(* IEC 61131-3 sources: plc-st-coding-agent/progress/evidence/f14_v10_full_20261113/jobs/custom_minimax-m27 (part 7) *)

(* ---- self-hard-04.raw_candidate_04.st ---- *)
FUNCTION_BLOCK FB
VAR_OUTPUT
    leadPump : INT := 0;
    lagPump : INT := 0;
    runningCount : INT := 0;
END_VAR
VAR_INPUT
    demand : INT;
    runHours : ARRAY[1..5] OF LINT;
    rotated : BOOL;
END_VAR
VAR
    tmp_prevLead : INT := 0;
    tmp_prevRunning : INT := 0;
    tmp_selectLag : BOOL := FALSE;
    tmp_newLead : INT;
    minHours : LINT;
    i : INT;
END_VAR
VAR_TEMP
    newLag : INT;
END_VAR
(*
ENGINEERING_CONTRACT:
  [S1] runningCount = CLAMP(demand, 0, 5). PUB001/PUB011
  [S2] demand=0→leadPump=lagPump=0; demand=1→lagPump=0; demand≥2→leadPump≠lagPump, both 1..5. PUB002/PUB012
  [S3] Lead-change requires old lead hours > new lead hours + 50. PUB036
  [S4] Hysteresis: rotated=TRUE AND runHours[lead] > minHours + 50 → rotate to min-hours pump. PUB026/PUB027
  [S5] Lag pump selected ONLY on: initial, lead change, runningCount increase. PUB005/PUB031
  [S6] Initial lead selection: min (runHours, pump#). PUB028
  [S7] Lag pump: min (runHours, pump#) excluding lead pump. PUB029
  [S8] Demand=0 clears lead/lag immediately; next positive demand triggers fresh selection. PUB033/PUB034
  [S9] First FB invocation initializes all outputs to 0 (VAR_INIT). PUB041
  No edge detection on rotated; it is level-triggered. PUB026
  Array bounds: 1..5 only. PUB042
*)
(* CONTRACT_RULES [] *)

tmp_prevLead := leadPump;
tmp_prevRunning := runningCount;
tmp_selectLag := FALSE;

minHours := runHours[1];
FOR i := 2 TO 5 DO
    IF runHours[i] < minHours THEN
        minHours := runHours[i];
    END_IF;
END_FOR;

IF demand <= 0 THEN
    runningCount := 0;
    leadPump := 0;
    lagPump := 0;
ELSIF leadPump = 0 THEN
    runningCount := demand;
    IF demand > 5 THEN
        runningCount := 5;
    ELSIF demand < 0 THEN
        runningCount := 0;
    END_IF;
    tmp_newLead := 1;
    FOR i := 2 TO 5 DO
        IF runHours[i] < runHours[tmp_newLead] OR (runHours[i] = runHours[tmp_newLead] AND i < tmp_newLead) THEN
            tmp_newLead := i;
        END_IF;
    END_FOR;
    leadPump := tmp_newLead;
    tmp_selectLag := TRUE;
    IF demand >= 2 THEN
        newLag := 0;
        FOR i := 1 TO 5 DO
            IF i <> leadPump THEN
                IF newLag = 0 OR runHours[i] < runHours[newLag] OR (runHours[i] = runHours[newLag] AND i < newLag) THEN
                    newLag := i;
                END_IF;
            END_IF;
        END_FOR;
        lagPump := newLag;
    ELSE
        lagPump := 0;
    END_IF;
ELSE
    IF demand > 5 THEN
        runningCount := 5;
    ELSIF demand < 0 THEN
        runningCount := 0;
    ELSE
        runningCount := demand;
    END_IF;
    IF rotated AND runHours[leadPump] > minHours + 50 THEN
        tmp_newLead := 1;
        FOR i := 2 TO 5 DO
            IF runHours[i] < runHours[tmp_newLead] OR (runHours[i] = runHours[tmp_newLead] AND i < tmp_newLead) THEN
                tmp_newLead := i;
            END_IF;
        END_FOR;
        leadPump := tmp_newLead;
        tmp_selectLag := TRUE;
    END_IF;
    IF demand > tmp_prevRunning THEN
        tmp_newLead := 1;
        FOR i := 2 TO 5 DO
            IF runHours[i] < runHours[tmp_newLead] OR (runHours[i] = runHours[tmp_newLead] AND i < tmp_newLead) THEN
                tmp_newLead := i;
            END_IF;
        END_FOR;
        leadPump := tmp_newLead;
        tmp_selectLag := TRUE;
    END_IF;
    IF tmp_selectLag THEN
        IF demand >= 2 THEN
            newLag := 0;
            FOR i := 1 TO 5 DO
                IF i <> leadPump THEN
                    IF newLag = 0 OR runHours[i] < runHours[newLag] OR (runHours[i] = runHours[newLag] AND i < newLag) THEN
                        newLag := i;
                    END_IF;
                END_IF;
            END_FOR;
            lagPump := newLag;
        ELSE
            lagPump := 0;
        END_IF;
    END_IF;
END_IF;
END_FUNCTION_BLOCK

(* ---- self-hard-05.candidate_01.st ---- *)
(* ENGINEERING_CONTRACT
 * FSM: Flame-trip latch with edge-reset.
 * [PUB001,PUB003] tripLatched activates SAME SCAN on (runRequest & !flameOK).
 * [PUB007] tripLatched holds until rising(resetBtn) & (!runRequest) & (!flameOK).
 *   Reset is edge-only; holding reset or pressing it under any other condition has no effect.
 * [PUB002,PUB004,PUB006] fuelPermit = runRequest & flameOK & !tripLatched (all three required).
 * [PUB005] o2Fault = !o2Valid OR o2PV<0 OR o2PV>21; fault removes trim only, never fuel.
 * [PUB008] trimEnable = fuelPermit & !o2Fault.
 * [PUB008,PUB030,PUB046] airTrim = 2.0*(2.0-o2PV) clamped [-10,+10]; 0 when trimEnable=FALSE.
 *   Positive limit never triggers (raw range [−38,+4] within o2PV∈[0,21]).
 * [PUB009,PUB031,PUB047] airCommand = baseAir+airTrim clamped [0,100]; 0 when fuelPermit=FALSE.
 *   baseAir may be outside [0,100]; final clamp applies to the sum only.
 *
 * LTL coverage:
 * S1  tripLatched on same-scan flame loss         → G((runRequest & !flameOK) → tripLatched)
 * S2  Self-hold; reset is edge-only               → G((prev(tripLatched) & !(rising & safe)) → tripLatched)
 * S3  tripLatched blocks fuel                     → G(tripLatched → !fuelPermit)
 * S4  fuelPermit full definition                  → G(fuelPermit ↔ runRequest & flameOK & !tripLatched)
 * S5  No fuel → airCommand=0                      → G(!fuelPermit → airCommand=0)
 * S6  airCommand ∈ [0,100]                        → G(airCommand≥0 ∧ airCommand≤100)
 * S7  airTrim ∈ [−10,10]                          → G(airTrim≥−10 ∧ airTrim≤10)
 * S8  trimEnable full definition                  → G(trimEnable ↔ fuelPermit & !o2Fault)
 * S9  o2Fault definition                          → G(o2Fault ↔ !o2Valid ∨ o2PV<0 ∨ o2PV>21)
 * S10 trimDisable → airTrim=0                     → G(!trimEnable → airTrim=0)
 * S11 o2PV>7 → negative clamp fires               → G((trimEnable & o2PV>7) → airTrim=−10)
 * S12 o2PV≤7 → no clamping                        → G((trimEnable & o2PV≤7) → airTrim=2*(2−o2PV))
 * S13 sum>100 → clamp to 100                      → G((fuelPermit & baseAir+airTrim>100) → airCommand=100)
 * S14 sum<0   → clamp to 0                        → G((fuelPermit & baseAir+airTrim<0)   → airCommand=0)
 * N10-S16 trip latch complete FSM                 → G(tripLatched ↔ (runRequest∧!flameOK)∨(prev∧!resetEdge)))
 * N10-S17 in-range sum is passed through          → G((fuelPermit & inRange) → airCommand=baseAir+airTrim)
 *
 * CONTRACT_RULES [{"kind":"hold_until_reset","output":"tripLatched","set_input":"runRequest","reset_input":"resetBtn"},{"kind":"hold_until_reset","output":"tripLatched","set_input":"flameOK","reset_input":"resetBtn"}]
 *)

FUNCTION_BLOCK FB
VAR_INPUT
    runRequest : BOOL;
    flameOK    : BOOL;
    o2Valid    : BOOL;
    o2PV       : REAL;
    baseAir    : REAL;
    resetBtn   : BOOL;
END_VAR
VAR_OUTPUT
    fuelPermit : BOOL;
    trimEnable : BOOL;
    airTrim    : REAL;
    airCommand : REAL;
    tripLatched: BOOL;
    o2Fault    : BOOL;
END_VAR
VAR
    prev_resetBtn   : BOOL := FALSE;
    prev_tripLatched: BOOL := FALSE;
END_VAR

    // --- Edge detection (same-scan memory) ---
    // Rising edge of resetBtn: was FALSE last scan, is TRUE this scan.
    // Store previous states at end of this scan for next invocation.

    // --- Flame-trip latch (PUB001,PUB003,PUB007) ---
    // Set on same scan when runRequest=TRUE and flameOK=FALSE.
    // Clear only on rising(resetBtn) AND runRequest=FALSE AND flameOK=FALSE.
    // Reset is edge-triggered; level-hold of resetBtn does NOT clear.
    IF runRequest AND NOT flameOK THEN
        tripLatched := TRUE;
    ELSIF prev_resetBtn = FALSE AND resetBtn = TRUE
          AND NOT runRequest AND NOT flameOK THEN
        tripLatched := FALSE;
    ELSE
        tripLatched := prev_tripLatched;
    END_IF;

    // --- Fuel permit (PUB002,PUB004,PUB006) ---
    fuelPermit := runRequest AND flameOK AND NOT tripLatched;

    // --- O2 fault detection (PUB005) ---
    o2Fault := NOT o2Valid OR o2PV < 0.0 OR o2PV > 21.0;

    // --- O2 trim correction (PUB008,PUB030,PUB046) ---
    trimEnable := fuelPermit AND NOT o2Fault;

    IF trimEnable THEN
        // Formula: 2.0 * (2.0 - o2PV), clamped to [-10, +10]
        // Within valid o2PV range [0,21] raw result lies in [-38, +4];
        // positive limit never triggers; negative limit fires when o2PV > 7.0.
        airTrim := 2.0 * (2.0 - o2PV);
        IF airTrim > 10.0 THEN
            airTrim := 10.0;
        ELSIF airTrim < -10.0 THEN
            airTrim := -10.0;
        END_IF;
    ELSE
        airTrim := 0.0;
    END_IF;

    // --- Air command (PUB009,PUB031,PUB047) ---
    // baseAir is external setpoint; may lie outside [0,100].
    // fuelPermit=FALSE forces airCommand to 0 (no residual position).
    IF fuelPermit THEN
        airCommand := baseAir + airTrim;
        IF airCommand > 100.0 THEN
            airCommand := 100.0;
        ELSIF airCommand < 0.0 THEN
            airCommand := 0.0;
        END_IF;
    ELSE
        airCommand := 0.0;
    END_IF;

    // --- Same-scan state update (persist for next scan) ---
    prev_resetBtn    := resetBtn;
    prev_tripLatched := tripLatched;
END_FUNCTION_BLOCK

(* ---- self-hard-05.raw_candidate_01.st ---- *)
(* ENGINEERING_CONTRACT
 * FSM: Flame-trip latch with edge-reset.
 * [PUB001,PUB003] tripLatched activates SAME SCAN on (runRequest & !flameOK).
 * [PUB007] tripLatched holds until rising(resetBtn) & (!runRequest) & (!flameOK).
 *   Reset is edge-only; holding reset or pressing it under any other condition has no effect.
 * [PUB002,PUB004,PUB006] fuelPermit = runRequest & flameOK & !tripLatched (all three required).
 * [PUB005] o2Fault = !o2Valid OR o2PV<0 OR o2PV>21; fault removes trim only, never fuel.
 * [PUB008] trimEnable = fuelPermit & !o2Fault.
 * [PUB008,PUB030,PUB046] airTrim = 2.0*(2.0-o2PV) clamped [-10,+10]; 0 when trimEnable=FALSE.
 *   Positive limit never triggers (raw range [−38,+4] within o2PV∈[0,21]).
 * [PUB009,PUB031,PUB047] airCommand = baseAir+airTrim clamped [0,100]; 0 when fuelPermit=FALSE.
 *   baseAir may be outside [0,100]; final clamp applies to the sum only.
 *
 * LTL coverage:
 * S1  tripLatched on same-scan flame loss         → G((runRequest & !flameOK) → tripLatched)
 * S2  Self-hold; reset is edge-only               → G((prev(tripLatched) & !(rising & safe)) → tripLatched)
 * S3  tripLatched blocks fuel                     → G(tripLatched → !fuelPermit)
 * S4  fuelPermit full definition                  → G(fuelPermit ↔ runRequest & flameOK & !tripLatched)
 * S5  No fuel → airCommand=0                      → G(!fuelPermit → airCommand=0)
 * S6  airCommand ∈ [0,100]                        → G(airCommand≥0 ∧ airCommand≤100)
 * S7  airTrim ∈ [−10,10]                          → G(airTrim≥−10 ∧ airTrim≤10)
 * S8  trimEnable full definition                  → G(trimEnable ↔ fuelPermit & !o2Fault)
 * S9  o2Fault definition                          → G(o2Fault ↔ !o2Valid ∨ o2PV<0 ∨ o2PV>21)
 * S10 trimDisable → airTrim=0                     → G(!trimEnable → airTrim=0)
 * S11 o2PV>7 → negative clamp fires               → G((trimEnable & o2PV>7) → airTrim=−10)
 * S12 o2PV≤7 → no clamping                        → G((trimEnable & o2PV≤7) → airTrim=2*(2−o2PV))
 * S13 sum>100 → clamp to 100                      → G((fuelPermit & baseAir+airTrim>100) → airCommand=100)
 * S14 sum<0   → clamp to 0                        → G((fuelPermit & baseAir+airTrim<0)   → airCommand=0)
 * N10-S16 trip latch complete FSM                 → G(tripLatched ↔ (runRequest∧!flameOK)∨(prev∧!resetEdge)))
 * N10-S17 in-range sum is passed through          → G((fuelPermit & inRange) → airCommand=baseAir+airTrim)
 *
 * CONTRACT_RULES [{"kind":"hold_until_reset","output":"tripLatched","set_input":"runRequest","reset_input":"resetBtn"},{"kind":"hold_until_reset","output":"tripLatched","set_input":"flameOK","reset_input":"resetBtn"}]
 *)

FUNCTION_BLOCK FB
VAR_INPUT
    runRequest : BOOL;
    flameOK    : BOOL;
    o2Valid    : BOOL;
    o2PV       : REAL;
    baseAir    : REAL;
    resetBtn   : BOOL;
END_VAR
VAR_OUTPUT
    fuelPermit : BOOL;
    trimEnable : BOOL;
    airTrim    : REAL;
    airCommand : REAL;
    tripLatched: BOOL;
    o2Fault    : BOOL;
END_VAR
VAR
    prev_resetBtn   : BOOL := FALSE;
    prev_tripLatched: BOOL := FALSE;
END_VAR

    // --- Edge detection (same-scan memory) ---
    // Rising edge of resetBtn: was FALSE last scan, is TRUE this scan.
    // Store previous states at end of this scan for next invocation.

    // --- Flame-trip latch (PUB001,PUB003,PUB007) ---
    // Set on same scan when runRequest=TRUE and flameOK=FALSE.
    // Clear only on rising(resetBtn) AND runRequest=FALSE AND flameOK=FALSE.
    // Reset is edge-triggered; level-hold of resetBtn does NOT clear.
    IF runRequest AND NOT flameOK THEN
        tripLatched := TRUE;
    ELSIF prev_resetBtn = FALSE AND resetBtn = TRUE
          AND NOT runRequest AND NOT flameOK THEN
        tripLatched := FALSE;
    ELSE
        tripLatched := prev_tripLatched;
    END_IF;

    // --- Fuel permit (PUB002,PUB004,PUB006) ---
    fuelPermit := runRequest AND flameOK AND NOT tripLatched;

    // --- O2 fault detection (PUB005) ---
    o2Fault := NOT o2Valid OR o2PV < 0.0 OR o2PV > 21.0;

    // --- O2 trim correction (PUB008,PUB030,PUB046) ---
    trimEnable := fuelPermit AND NOT o2Fault;

    IF trimEnable THEN
        // Formula: 2.0 * (2.0 - o2PV), clamped to [-10, +10]
        // Within valid o2PV range [0,21] raw result lies in [-38, +4];
        // positive limit never triggers; negative limit fires when o2PV > 7.0.
        airTrim := 2.0 * (2.0 - o2PV);
        IF airTrim > 10.0 THEN
            airTrim := 10.0;
        ELSIF airTrim < -10.0 THEN
            airTrim := -10.0;
        END_IF;
    ELSE
        airTrim := 0.0;
    END_IF;

    // --- Air command (PUB009,PUB031,PUB047) ---
    // baseAir is external setpoint; may lie outside [0,100].
    // fuelPermit=FALSE forces airCommand to 0 (no residual position).
    IF fuelPermit THEN
        airCommand := baseAir + airTrim;
        IF airCommand > 100.0 THEN
            airCommand := 100.0;
        ELSIF airCommand < 0.0 THEN
            airCommand := 0.0;
        END_IF;
    ELSE
        airCommand := 0.0;
    END_IF;

    // --- Same-scan state update (persist for next scan) ---
    prev_resetBtn    := resetBtn;
    prev_tripLatched := tripLatched;
END_FUNCTION_BLOCK

(* ---- self-hard-06.candidate_01.st ---- *)
(* CONTRACT_RULES [{"kind": "hold_until_reset", "output": "tripLatched", "set_input": "runRequest_AND_NOT_pressureValid_OR_pressure_ge_4500", "reset_input": "resetBtn_rising_AND_NOT_runRequest_AND_pressureValid_AND_pressure_le_4200"}] *)
(* ENGINEERING_CONTRACT
   PUB001-PUB004:  Trip activation same-scan when runRequest AND (NOT pressureValid OR pressure >= 4500.0 kPa).
   PUB005:         Hysteresis band 300 kPa: reset clears only when pressure <= 4200.0 (strict <=).
   PUB006-PUB008:  tripLatched holds until resetBtn rising edge + NOT runRequest + pressureValid + pressure <= 4200.0.
   PUB009-PUB011:  currentCauseMask LOW-4 encoding: bit0=xmitter fail, bit1=valve stick(3-consecutive), bit2=excess combustion, bit3=unlocated.
                    Only evaluated when runRequest AND pressureValid AND pressure >= 4500.0 (bits 1/2); bit0 when runRequest AND NOT pressureValid.
                    Not runRequest → mask = 0.
   PUB012-PUB014:  Valve stick counter requires 3 consecutive cycles of (runRequest AND pressureValid AND pressure >= 4500.0 AND outletCmd >= 50 AND outletFeedback <= 10).
                    Any break (feedback OK, pressure < 4500, pressureValid=FALSE, runRequest=FALSE) → counter = 0.
   PUB015-PUB017:  latchedCauseMask accumulates via bitwise OR each scan tripLatched is TRUE (16-bit WORD, max 15, no overflow).
                    Cleared only on legal reset. Reflects full trip history, not a snapshot.
   PUB018-PUB020:  fuelPermit = runRequest AND NOT tripLatched; diagnosticActive = (currentCauseMask <> 0).
   PUB021-PUB023:  Clue encodings: 0=none, 1=xmitter fail, 2=stick only, 4=combustion only, 6=both, 8=unlocated.
   Units: kPa (pressure), t/h (flow), % (valve), ms TON timers (not used; discrete-cycle counting).
*)
FUNCTION_BLOCK FB
VAR
    prevResetBtn      : BOOL := FALSE;   // PUB006: previous scan resetBtn for R_TRIG
    prevStickingCond1 : BOOL := FALSE;   // N10-S11: condition state at scan N-1
    prevStickingCond2 : BOOL := FALSE;   // N10-S11: condition state at scan N-2
    stickingCount     : INT  := 0;       // PUB012: consecutive-cycle counter (0..3)
END_VAR
VAR_OUTPUT
    tripLatched       : BOOL;
    fuelPermit        : BOOL;
    currentCauseMask  : WORD;
    latchedCauseMask  : WORD;
    diagnosticActive  : BOOL;
END_VAR

    // --- Rising-edge detection for reset button (PUB006) ---
    VAR temp_resetRising : BOOL;
    temp_resetRising := resetBtn AND NOT prevResetBtn;

    // --- Trip condition (PUB001-PUB004, S1, S2, S17) ---
    // Set: runRequest AND (NOT pressureValid OR pressure >= 4500.0)
    // Clear: rising resetBtn AND NOT runRequest AND pressureValid AND pressure <= 4200.0
    IF temp_resetRising AND NOT runRequest AND pressureValid AND (pressure <= 4200.0) THEN
        tripLatched := FALSE;
    ELSIF runRequest AND (NOT pressureValid OR (pressure >= 4500.0)) THEN
        tripLatched := TRUE;
    END_IF;

    // --- Valve sticking: 3 consecutive cycles under valid overpressure (PUB012-PUB014, N10-S11) ---
    // Condition: runRequest AND pressureValid AND pressure >= 4500.0 AND outletCmd >= 50 AND outletFeedback <= 10
    IF runRequest AND pressureValid AND (pressure >= 4500.0) AND (outletCmd >= 50) AND (outletFeedback <= 10) THEN
        // All three cycles met: current + prev1 + prev2
        IF prevStickingCond1 AND prevStickingCond2 THEN
            stickingCount := 3;
        ELSE
            stickingCount := stickingCount + 1;
            IF stickingCount > 3 THEN
                stickingCount := 3;
            END_IF;
        END_IF;
    ELSE
        // Any break resets counter (PUB014: feedback OK / pressure drop / invalid / stop)
        stickingCount := 0;
    END_IF;

    // --- Current cause mask (PUB009-PUB011, S5, S6, S9-S12, N10-S10, N10-S11, N10-S15) ---
    currentCauseMask := 16#0000;

    IF NOT runRequest THEN
        // PUB009: Not runRequest → mask = 0
        currentCauseMask := 16#0000;
    ELSIF NOT pressureValid THEN
        // PUB010: bit0=1 Transmitter failure (worst-case trip, PUB001)
        currentCauseMask := 16#0001;
    ELSE
        // pressureValid = TRUE
        IF pressure >= 4500.0 THEN
            // Evaluate bit1 (valve sticking) and bit2 (excess combustion) only in overpressure工况 (PUB010)
            // bit1: 3 consecutive cycles
            IF stickingCount >= 3 THEN
                currentCauseMask := currentCauseMask OR INT_TO_WORD(2); // bit1=2
            END_IF;

            // bit2: Excess combustion
            IF (fuelFlow >= 4.0) AND (steamFlow <= 10.0) THEN
                currentCauseMask := currentCauseMask OR INT_TO_WORD(4); // bit2=4
            END_IF;

            // bit3=8: Unlocated (overpressure but neither bit1 nor bit2 set, PUB010)
            IF (stickingCount < 3) AND NOT ((fuelFlow >= 4.0) AND (steamFlow <= 10.0)) THEN
                currentCauseMask := currentCauseMask OR INT_TO_WORD(8); // bit3=8
            END_IF;
        END_IF;
        // pressure < 4500.0: no clues (S6, N10-S15)
    END_IF;

    // --- Latched cause mask accumulation (PUB015-PUB017, S13, N10-S18) ---
    // Accumulates full trip history via bitwise OR while tripLatched is TRUE
    IF tripLatched AND (currentCauseMask <> 16#0000) THEN
        latchedCauseMask := latchedCauseMask OR currentCauseMask;
    END_IF;

    // --- Outputs (PUB018-PUB020, S3, N10-S16) ---
    fuelPermit       := runRequest AND NOT tripLatched;
    diagnosticActive := (currentCauseMask <> 16#0000);

    // --- State propagation for next scan ---
    prevResetBtn      := resetBtn;
    prevStickingCond2 := prevStickingCond1;
    prevStickingCond1 := (runRequest AND pressureValid AND (pressure >= 4500.0) AND (outletCmd >= 50) AND (outletFeedback <= 10));

END_FUNCTION_BLOCK

(* ---- self-hard-06.candidate_02.st ---- *)
(* CONTRACT_RULES [{"kind": "hold_until_reset", "output": "tripLatched", "set_input": "runRequest_AND_NOT_pressureValid_OR_pressure_ge_4500", "reset_input": "resetBtn_rising_AND_NOT_runRequest_AND_pressureValid_AND_pressure_le_4200"}] *)
(* ENGINEERING_CONTRACT
   PUB001-PUB004:  Trip activation same-scan when runRequest AND (NOT pressureValid OR pressure >= 4500.0 kPa).
   PUB005:         Hysteresis band 300 kPa: reset clears only when pressure <= 4200.0 (strict <=).
   PUB006-PUB008:  tripLatched holds until resetBtn rising edge + NOT runRequest + pressureValid + pressure <= 4200.0.
   PUB009-PUB011:  currentCauseMask LOW-4 encoding: bit0=xmitter fail, bit1=valve stick(3-consecutive), bit2=excess combustion, bit3=unlocated.
                    Only evaluated when runRequest AND pressureValid AND pressure >= 4500.0 (bits 1/2); bit0 when runRequest AND NOT pressureValid.
                    Not runRequest → mask = 0.
   PUB012-PUB014:  Valve stick counter requires 3 consecutive cycles of (runRequest AND pressureValid AND pressure >= 4500.0 AND outletCmd >= 50 AND outletFeedback <= 10).
                    Any break (feedback OK, pressure < 4500, pressureValid=FALSE, runRequest=FALSE) → counter = 0.
   PUB015-PUB017:  latchedCauseMask accumulates via bitwise OR each scan tripLatched is TRUE (16-bit WORD, max 15, no overflow).
                    Cleared only on legal reset. Reflects full trip history, not a snapshot.
   PUB018-PUB020:  fuelPermit = runRequest AND NOT tripLatched; diagnosticActive = (currentCauseMask <> 0).
   PUB021-PUB023:  Clue encodings: 0=none, 1=xmitter fail, 2=stick only, 4=combustion only, 6=both, 8=unlocated.
   Units: kPa (pressure), t/h (flow), % (valve), ms TON timers (not used; discrete-cycle counting).
*)
FUNCTION_BLOCK FB
VAR
    prevResetBtn      : BOOL := FALSE;
    prevStickingCond1 : BOOL := FALSE;
    prevStickingCond2 : BOOL := FALSE;
    stickingCount     : INT  := 0;
    tempResetRising   : BOOL := FALSE;
END_VAR
VAR_OUTPUT
    tripLatched       : BOOL;
    fuelPermit        : BOOL;
    currentCauseMask  : WORD;
    latchedCauseMask  : WORD;
    diagnosticActive  : BOOL;
END_VAR

    // --- Rising-edge detection for reset button (PUB006) ---
    tempResetRising := resetBtn AND NOT prevResetBtn;

    // --- Trip condition (PUB001-PUB004, S1, S2, S17) ---
    IF tempResetRising AND NOT runRequest AND pressureValid AND (pressure <= 4200.0) THEN
        tripLatched := FALSE;
    ELSIF runRequest AND (NOT pressureValid OR (pressure >= 4500.0)) THEN
        tripLatched := TRUE;
    END_IF;

    // --- Valve sticking: 3 consecutive cycles under valid overpressure (PUB012-PUB014, N10-S11) ---
    IF runRequest AND pressureValid AND (pressure >= 4500.0) AND (outletCmd >= 50) AND (outletFeedback <= 10) THEN
        IF prevStickingCond1 AND prevStickingCond2 THEN
            stickingCount := 3;
        ELSE
            stickingCount := stickingCount + 1;
            IF stickingCount > 3 THEN
                stickingCount := 3;
            END_IF;
        END_IF;
    ELSE
        stickingCount := 0;
    END_IF;

    // --- Current cause mask (PUB009-PUB011, S5, S6, S9-S12, N10-S10, N10-S11, N10-S15) ---
    currentCauseMask := 16#0000;

    IF NOT runRequest THEN
        currentCauseMask := 16#0000;
    ELSIF NOT pressureValid THEN
        currentCauseMask := 16#0001;
    ELSE
        IF pressure >= 4500.0 THEN
            IF stickingCount >= 3 THEN
                currentCauseMask := currentCauseMask OR TO_WORD(2);
            END_IF;
            IF (fuelFlow >= 4.0) AND (steamFlow <= 10.0) THEN
                currentCauseMask := currentCauseMask OR TO_WORD(4);
            END_IF;
            IF (stickingCount < 3) AND NOT ((fuelFlow >= 4.0) AND (steamFlow <= 10.0)) THEN
                currentCauseMask := currentCauseMask OR TO_WORD(8);
            END_IF;
        END_IF;
    END_IF;

    // --- Latched cause mask accumulation (PUB015-PUB017, S13, N10-S18) ---
    IF tripLatched AND (currentCauseMask <> 16#0000) THEN
        latchedCauseMask := latchedCauseMask OR currentCauseMask;
    END_IF;

    // --- Outputs (PUB018-PUB020, S3, N10-S16) ---
    fuelPermit       := runRequest AND NOT tripLatched;
    diagnosticActive := (currentCauseMask <> 16#0000);

    // --- State propagation for next scan ---
    prevResetBtn      := resetBtn;
    prevStickingCond2 := prevStickingCond1;
    prevStickingCond1 := (runRequest AND pressureValid AND (pressure >= 4500.0) AND (outletCmd >= 50) AND (outletFeedback <= 10));

END_FUNCTION_BLOCK

(* ---- self-hard-06.candidate_03.st ---- *)
(* CONTRACT_RULES [{"kind": "hold_until_reset", "output": "tripLatched", "set_input": "runRequest_AND_NOT_pressureValid_OR_pressure_ge_4500", "reset_input": "resetBtn_rising_AND_NOT_runRequest_AND_pressureValid_AND_pressure_le_4200"}] *)
(* ENGINEERING_CONTRACT
   PUB001-PUB004:  Trip activation same-scan when runRequest AND (NOT pressureValid OR pressure >= 4500.0 kPa).
   PUB005:         Hysteresis band 300 kPa: reset clears only when pressure <= 4200.0 (strict <=).
   PUB006-PUB008:  tripLatched holds until resetBtn rising edge + NOT runRequest + pressureValid + pressure <= 4200.0.
   PUB009-PUB011:  currentCauseMask LOW-4 encoding: bit0=xmitter fail, bit1=valve stick(3-consecutive), bit2=excess combustion, bit3=unlocated.
                    Only evaluated when runRequest AND pressureValid AND pressure >= 4500.0 (bits 1/2); bit0 when runRequest AND NOT pressureValid.
                    Not runRequest → mask = 0.
   PUB012-PUB014:  Valve stick counter requires 3 consecutive cycles of (runRequest AND pressureValid AND pressure >= 4500.0 AND outletCmd >= 50 AND outletFeedback <= 10).
                    Any break (feedback OK, pressure < 4500, pressureValid=FALSE, runRequest=FALSE) → counter = 0.
   PUB015-PUB017:  latchedCauseMask accumulates via bitwise OR each scan tripLatched is TRUE (16-bit WORD, max 15, no overflow).
                    Cleared only on legal reset. Reflects full trip history, not a snapshot.
   PUB018-PUB020:  fuelPermit = runRequest AND NOT tripLatched; diagnosticActive = (currentCauseMask <> 0).
   PUB021-PUB023:  Clue encodings: 0=none, 1=xmitter fail, 2=stick only, 4=combustion only, 6=both, 8=unlocated.
   Units: kPa (pressure), t/h (flow), % (valve).
*)
FUNCTION_BLOCK FB
VAR
    prevResetBtn      : BOOL := FALSE;
    prevStickingCond1 : BOOL := FALSE;
    prevStickingCond2 : BOOL := FALSE;
    stickingCount     : INT  := 0;
    local_tripLatched : BOOL := FALSE;
    local_fuelPermit  : BOOL := FALSE;
    local_currentMask : WORD := 16#0000;
    local_latchedMask : WORD := 16#0000;
END_VAR
VAR_TEMP
    resetRising   : BOOL;
    curSticking   : BOOL;
END_VAR

    resetRising := resetBtn AND NOT prevResetBtn;

    IF resetRising AND NOT runRequest AND pressureValid AND (pressure <= 4200.0) THEN
        local_tripLatched := FALSE;
        local_latchedMask := 16#0000;
    ELSIF runRequest AND (NOT pressureValid OR (pressure >= 4500.0)) THEN
        local_tripLatched := TRUE;
    END_IF;

    curSticking := runRequest AND pressureValid AND (pressure >= 4500.0) AND (outletCmd >= 50) AND (outletFeedback <= 10);

    IF curSticking THEN
        IF prevStickingCond1 AND prevStickingCond2 THEN
            stickingCount := 3;
        ELSE
            stickingCount := stickingCount + 1;
            IF stickingCount > 3 THEN
                stickingCount := 3;
            END_IF;
        END_IF;
    ELSE
        stickingCount := 0;
    END_IF;

    local_currentMask := 16#0000;

    IF NOT runRequest THEN
        local_currentMask := 16#0000;
    ELSIF NOT pressureValid THEN
        local_currentMask := 16#0001;
    ELSE
        IF pressure >= 4500.0 THEN
            IF stickingCount >= 3 THEN
                local_currentMask := local_currentMask OR TO_WORD(2);
            END_IF;
            IF (fuelFlow >= 4.0) AND (steamFlow <= 10.0) THEN
                local_currentMask := local_currentMask OR TO_WORD(4);
            END_IF;
            IF (stickingCount < 3) AND NOT ((fuelFlow >= 4.0) AND (steamFlow <= 10.0)) THEN
                local_currentMask := local_currentMask OR TO_WORD(8);
            END_IF;
        END_IF;
    END_IF;

    IF local_tripLatched THEN
        local_latchedMask := local_latchedMask OR local_currentMask;
    END_IF;

    local_fuelPermit := runRequest AND NOT local_tripLatched;

    tripLatched      := local_tripLatched;
    fuelPermit       := local_fuelPermit;
    currentCauseMask := local_currentMask;
    latchedCauseMask := local_latchedMask;
    diagnosticActive := (local_currentMask <> 16#0000);

    prevResetBtn      := resetBtn;
    prevStickingCond2 := prevStickingCond1;
    prevStickingCond1 := curSticking;

END_FUNCTION_BLOCK

(* ---- self-hard-06.candidate_04.st ---- *)
(* CONTRACT_RULES [{"kind": "hold_until_reset", "output": "tripLatched", "set_input": "runRequest_AND_NOT_pressureValid_OR_pressure_ge_4500", "reset_input": "resetBtn_rising_AND_NOT_runRequest_AND_pressureValid_AND_pressure_le_4200"}] *)
(* ENGINEERING_CONTRACT
   PUB001-PUB004:  Trip activation same-scan when runRequest AND (NOT pressureValid OR pressure >= 4500.0 kPa).
   PUB005:         Hysteresis band 300 kPa: reset clears only when pressure <= 4200.0 (strict <=).
   PUB006-PUB008:  tripLatched holds until resetBtn rising edge + NOT runRequest + pressureValid + pressure <= 4200.0.
   PUB009-PUB011:  currentCauseMask LOW-4 encoding: bit0=xmitter fail, bit1=valve stick(3-consecutive), bit2=excess combustion, bit3=unlocated.
                    Only evaluated when runRequest AND pressureValid AND pressure >= 4500.0 (bits 1/2); bit0 when runRequest AND NOT pressureValid.
                    Not runRequest → mask = 0.
   PUB012-PUB014:  Valve stick counter requires 3 consecutive cycles of (runRequest AND pressureValid AND pressure >= 4500.0 AND outletCmd >= 50 AND outletFeedback <= 10).
                    Any break (feedback OK, pressure < 4500, pressureValid=FALSE, runRequest=FALSE) → counter = 0.
   PUB015-PUB017:  latchedCauseMask accumulates via bitwise OR each scan tripLatched is TRUE (16-bit WORD, max 15, no overflow).
                    Cleared only on legal reset. Reflects full trip history, not a snapshot.
   PUB018-PUB020:  fuelPermit = runRequest AND NOT tripLatched; diagnosticActive = (currentCauseMask <> 0).
   PUB021-PUB023:  Clue encodings: 0=none, 1=xmitter fail, 2=stick only, 4=combustion only, 6=both, 8=unlocated.
   Units: kPa (pressure), t/h (flow), % (valve).
*)
FUNCTION_BLOCK FB
VAR
    prevResetBtn      : BOOL := FALSE;
    prevStickingCond1 : BOOL := FALSE;
    prevStickingCond2 : BOOL := FALSE;
    stickingCount     : INT  := 0;
    tmpResetRising    : BOOL := FALSE;
END_VAR
VAR_OUTPUT
    tripLatched       : BOOL;
    fuelPermit        : BOOL;
    currentCauseMask  : WORD;
    latchedCauseMask  : WORD;
    diagnosticActive  : BOOL;
END_VAR

    // Rising-edge detection for reset button (PUB006)
    tmpResetRising := resetBtn AND NOT prevResetBtn;

    // Trip condition: set or clear tripLatched (PUB001-PUB004, S1, S2, S17)
    IF tmpResetRising AND NOT runRequest AND pressureValid AND (pressure <= 4200.0) THEN
        tripLatched := FALSE;
    ELSIF runRequest AND (NOT pressureValid OR (pressure >= 4500.0)) THEN
        tripLatched := TRUE;
    END_IF;

    // Valve sticking: 3 consecutive cycles under valid overpressure (PUB012-PUB014, N10-S11)
    IF runRequest AND pressureValid AND (pressure >= 4500.0) AND (outletCmd >= 50) AND (outletFeedback <= 10) THEN
        IF prevStickingCond1 AND prevStickingCond2 THEN
            stickingCount := 3;
        ELSE
            stickingCount := stickingCount + 1;
            IF stickingCount > 3 THEN
                stickingCount := 3;
            END_IF;
        END_IF;
    ELSE
        stickingCount := 0;
    END_IF;

    // Current cause mask (PUB009-PUB011, S5, S6, S9-S12, N10-S10, N10-S11, N10-S15)
    currentCauseMask := 16#0000;

    IF NOT runRequest THEN
        currentCauseMask := 16#0000;
    ELSIF NOT pressureValid THEN
        currentCauseMask := 16#0001;
    ELSE
        IF pressure >= 4500.0 THEN
            IF stickingCount >= 3 THEN
                currentCauseMask := currentCauseMask OR INT_TO_WORD(2);
            END_IF;
            IF (fuelFlow >= 4.0) AND (steamFlow <= 10.0) THEN
                currentCauseMask := currentCauseMask OR INT_TO_WORD(4);
            END_IF;
            IF (stickingCount < 3) AND NOT ((fuelFlow >= 4.0) AND (steamFlow <= 10.0)) THEN
                currentCauseMask := currentCauseMask OR INT_TO_WORD(8);
            END_IF;
        END_IF;
    END_IF;

    // Latched cause mask accumulation (PUB015-PUB017, S13, N10-S18)
    IF tripLatched AND (currentCauseMask <> 16#0000) THEN
        latchedCauseMask := latchedCauseMask OR currentCauseMask;
    END_IF;

    // Outputs (PUB018-PUB020, S3, N10-S16)
    fuelPermit       := runRequest AND NOT tripLatched;
    diagnosticActive := (currentCauseMask <> 16#0000);

    // State propagation for next scan
    prevResetBtn      := resetBtn;
    prevStickingCond2 := prevStickingCond1;
    prevStickingCond1 := (runRequest AND pressureValid AND (pressure >= 4500.0) AND (outletCmd >= 50) AND (outletFeedback <= 10));

END_FUNCTION_BLOCK

(* ---- self-hard-06.raw_candidate_01.st ---- *)
(* CONTRACT_RULES [{"kind": "hold_until_reset", "output": "tripLatched", "set_input": "runRequest_AND_NOT_pressureValid_OR_pressure_ge_4500", "reset_input": "resetBtn_rising_AND_NOT_runRequest_AND_pressureValid_AND_pressure_le_4200"}] *)
(* ENGINEERING_CONTRACT
   PUB001-PUB004:  Trip activation same-scan when runRequest AND (NOT pressureValid OR pressure >= 4500.0 kPa).
   PUB005:         Hysteresis band 300 kPa: reset clears only when pressure <= 4200.0 (strict <=).
   PUB006-PUB008:  tripLatched holds until resetBtn rising edge + NOT runRequest + pressureValid + pressure <= 4200.0.
   PUB009-PUB011:  currentCauseMask LOW-4 encoding: bit0=xmitter fail, bit1=valve stick(3-consecutive), bit2=excess combustion, bit3=unlocated.
                    Only evaluated when runRequest AND pressureValid AND pressure >= 4500.0 (bits 1/2); bit0 when runRequest AND NOT pressureValid.
                    Not runRequest → mask = 0.
   PUB012-PUB014:  Valve stick counter requires 3 consecutive cycles of (runRequest AND pressureValid AND pressure >= 4500.0 AND outletCmd >= 50 AND outletFeedback <= 10).
                    Any break (feedback OK, pressure < 4500, pressureValid=FALSE, runRequest=FALSE) → counter = 0.
   PUB015-PUB017:  latchedCauseMask accumulates via bitwise OR each scan tripLatched is TRUE (16-bit WORD, max 15, no overflow).
                    Cleared only on legal reset. Reflects full trip history, not a snapshot.
   PUB018-PUB020:  fuelPermit = runRequest AND NOT tripLatched; diagnosticActive = (currentCauseMask <> 0).
   PUB021-PUB023:  Clue encodings: 0=none, 1=xmitter fail, 2=stick only, 4=combustion only, 6=both, 8=unlocated.
   Units: kPa (pressure), t/h (flow), % (valve), ms TON timers (not used; discrete-cycle counting).
*)
FUNCTION_BLOCK FB
VAR
    prevResetBtn      : BOOL := FALSE;   // PUB006: previous scan resetBtn for R_TRIG
    prevStickingCond1 : BOOL := FALSE;   // N10-S11: condition state at scan N-1
    prevStickingCond2 : BOOL := FALSE;   // N10-S11: condition state at scan N-2
    stickingCount     : INT  := 0;       // PUB012: consecutive-cycle counter (0..3)
END_VAR
VAR_OUTPUT
    tripLatched       : BOOL;
    fuelPermit        : BOOL;
    currentCauseMask  : WORD;
    latchedCauseMask  : WORD;
    diagnosticActive  : BOOL;
END_VAR

    // --- Rising-edge detection for reset button (PUB006) ---
    VAR temp_resetRising : BOOL;
    temp_resetRising := resetBtn AND NOT prevResetBtn;

    // --- Trip condition (PUB001-PUB004, S1, S2, S17) ---
    // Set: runRequest AND (NOT pressureValid OR pressure >= 4500.0)
    // Clear: rising resetBtn AND NOT runRequest AND pressureValid AND pressure <= 4200.0
    IF temp_resetRising AND NOT runRequest AND pressureValid AND (pressure <= 4200.0) THEN
        tripLatched := FALSE;
    ELSIF runRequest AND (NOT pressureValid OR (pressure >= 4500.0)) THEN
        tripLatched := TRUE;
    END_IF;

    // --- Valve sticking: 3 consecutive cycles under valid overpressure (PUB012-PUB014, N10-S11) ---
    // Condition: runRequest AND pressureValid AND pressure >= 4500.0 AND outletCmd >= 50 AND outletFeedback <= 10
    IF runRequest AND pressureValid AND (pressure >= 4500.0) AND (outletCmd >= 50) AND (outletFeedback <= 10) THEN
        // All three cycles met: current + prev1 + prev2
        IF prevStickingCond1 AND prevStickingCond2 THEN
            stickingCount := 3;
        ELSE
            stickingCount := stickingCount + 1;
            IF stickingCount > 3 THEN
                stickingCount := 3;
            END_IF;
        END_IF;
    ELSE
        // Any break resets counter (PUB014: feedback OK / pressure drop / invalid / stop)
        stickingCount := 0;
    END_IF;

    // --- Current cause mask (PUB009-PUB011, S5, S6, S9-S12, N10-S10, N10-S11, N10-S15) ---
    currentCauseMask := 16#0000;

    IF NOT runRequest THEN
        // PUB009: Not runRequest → mask = 0
        currentCauseMask := 16#0000;
    ELSIF NOT pressureValid THEN
        // PUB010: bit0=1 Transmitter failure (worst-case trip, PUB001)
        currentCauseMask := 16#0001;
    ELSE
        // pressureValid = TRUE
        IF pressure >= 4500.0 THEN
            // Evaluate bit1 (valve sticking) and bit2 (excess combustion) only in overpressure工况 (PUB010)
            // bit1: 3 consecutive cycles
            IF stickingCount >= 3 THEN
                currentCauseMask := currentCauseMask OR INT_TO_WORD(2); // bit1=2
            END_IF;

            // bit2: Excess combustion
            IF (fuelFlow >= 4.0) AND (steamFlow <= 10.0) THEN
                currentCauseMask := currentCauseMask OR INT_TO_WORD(4); // bit2=4
            END_IF;

            // bit3=8: Unlocated (overpressure but neither bit1 nor bit2 set, PUB010)
            IF (stickingCount < 3) AND NOT ((fuelFlow >= 4.0) AND (steamFlow <= 10.0)) THEN
                currentCauseMask := currentCauseMask OR INT_TO_WORD(8); // bit3=8
            END_IF;
        END_IF;
        // pressure < 4500.0: no clues (S6, N10-S15)
    END_IF;

    // --- Latched cause mask accumulation (PUB015-PUB017, S13, N10-S18) ---
    // Accumulates full trip history via bitwise OR while tripLatched is TRUE
    IF tripLatched AND (currentCauseMask <> 16#0000) THEN
        latchedCauseMask := latchedCauseMask OR currentCauseMask;
    END_IF;

    // --- Outputs (PUB018-PUB020, S3, N10-S16) ---
    fuelPermit       := runRequest AND NOT tripLatched;
    diagnosticActive := (currentCauseMask <> 16#0000);

    // --- State propagation for next scan ---
    prevResetBtn      := resetBtn;
    prevStickingCond2 := prevStickingCond1;
    prevStickingCond1 := (runRequest AND pressureValid AND (pressure >= 4500.0) AND (outletCmd >= 50) AND (outletFeedback <= 10));

END_FUNCTION_BLOCK

(* ---- self-hard-06.raw_candidate_02.st ---- *)
(* CONTRACT_RULES [{"kind": "hold_until_reset", "output": "tripLatched", "set_input": "runRequest_AND_NOT_pressureValid_OR_pressure_ge_4500", "reset_input": "resetBtn_rising_AND_NOT_runRequest_AND_pressureValid_AND_pressure_le_4200"}] *)
(* ENGINEERING_CONTRACT
   PUB001-PUB004:  Trip activation same-scan when runRequest AND (NOT pressureValid OR pressure >= 4500.0 kPa).
   PUB005:         Hysteresis band 300 kPa: reset clears only when pressure <= 4200.0 (strict <=).
   PUB006-PUB008:  tripLatched holds until resetBtn rising edge + NOT runRequest + pressureValid + pressure <= 4200.0.
   PUB009-PUB011:  currentCauseMask LOW-4 encoding: bit0=xmitter fail, bit1=valve stick(3-consecutive), bit2=excess combustion, bit3=unlocated.
                    Only evaluated when runRequest AND pressureValid AND pressure >= 4500.0 (bits 1/2); bit0 when runRequest AND NOT pressureValid.
                    Not runRequest → mask = 0.
   PUB012-PUB014:  Valve stick counter requires 3 consecutive cycles of (runRequest AND pressureValid AND pressure >= 4500.0 AND outletCmd >= 50 AND outletFeedback <= 10).
                    Any break (feedback OK, pressure < 4500, pressureValid=FALSE, runRequest=FALSE) → counter = 0.
   PUB015-PUB017:  latchedCauseMask accumulates via bitwise OR each scan tripLatched is TRUE (16-bit WORD, max 15, no overflow).
                    Cleared only on legal reset. Reflects full trip history, not a snapshot.
   PUB018-PUB020:  fuelPermit = runRequest AND NOT tripLatched; diagnosticActive = (currentCauseMask <> 0).
   PUB021-PUB023:  Clue encodings: 0=none, 1=xmitter fail, 2=stick only, 4=combustion only, 6=both, 8=unlocated.
   Units: kPa (pressure), t/h (flow), % (valve), ms TON timers (not used; discrete-cycle counting).
*)
FUNCTION_BLOCK FB
VAR
    prevResetBtn      : BOOL := FALSE;
    prevStickingCond1 : BOOL := FALSE;
    prevStickingCond2 : BOOL := FALSE;
    stickingCount     : INT  := 0;
    tempResetRising   : BOOL := FALSE;
END_VAR
VAR_OUTPUT
    tripLatched       : BOOL;
    fuelPermit        : BOOL;
    currentCauseMask  : WORD;
    latchedCauseMask  : WORD;
    diagnosticActive  : BOOL;
END_VAR

    // --- Rising-edge detection for reset button (PUB006) ---
    tempResetRising := resetBtn AND NOT prevResetBtn;

    // --- Trip condition (PUB001-PUB004, S1, S2, S17) ---
    IF tempResetRising AND NOT runRequest AND pressureValid AND (pressure <= 4200.0) THEN
        tripLatched := FALSE;
    ELSIF runRequest AND (NOT pressureValid OR (pressure >= 4500.0)) THEN
        tripLatched := TRUE;
    END_IF;

    // --- Valve sticking: 3 consecutive cycles under valid overpressure (PUB012-PUB014, N10-S11) ---
    IF runRequest AND pressureValid AND (pressure >= 4500.0) AND (outletCmd >= 50) AND (outletFeedback <= 10) THEN
        IF prevStickingCond1 AND prevStickingCond2 THEN
            stickingCount := 3;
        ELSE
            stickingCount := stickingCount + 1;
            IF stickingCount > 3 THEN
                stickingCount := 3;
            END_IF;
        END_IF;
    ELSE
        stickingCount := 0;
    END_IF;

    // --- Current cause mask (PUB009-PUB011, S5, S6, S9-S12, N10-S10, N10-S11, N10-S15) ---
    currentCauseMask := 16#0000;

    IF NOT runRequest THEN
        currentCauseMask := 16#0000;
    ELSIF NOT pressureValid THEN
        currentCauseMask := 16#0001;
    ELSE
        IF pressure >= 4500.0 THEN
            IF stickingCount >= 3 THEN
                currentCauseMask := currentCauseMask OR TO_WORD(2);
            END_IF;
            IF (fuelFlow >= 4.0) AND (steamFlow <= 10.0) THEN
                currentCauseMask := currentCauseMask OR TO_WORD(4);
            END_IF;
            IF (stickingCount < 3) AND NOT ((fuelFlow >= 4.0) AND (steamFlow <= 10.0)) THEN
                currentCauseMask := currentCauseMask OR TO_WORD(8);
            END_IF;
        END_IF;
    END_IF;

    // --- Latched cause mask accumulation (PUB015-PUB017, S13, N10-S18) ---
    IF tripLatched AND (currentCauseMask <> 16#0000) THEN
        latchedCauseMask := latchedCauseMask OR currentCauseMask;
    END_IF;

    // --- Outputs (PUB018-PUB020, S3, N10-S16) ---
    fuelPermit       := runRequest AND NOT tripLatched;
    diagnosticActive := (currentCauseMask <> 16#0000);

    // --- State propagation for next scan ---
    prevResetBtn      := resetBtn;
    prevStickingCond2 := prevStickingCond1;
    prevStickingCond1 := (runRequest AND pressureValid AND (pressure >= 4500.0) AND (outletCmd >= 50) AND (outletFeedback <= 10));

END_FUNCTION_BLOCK

(* ---- self-hard-06.raw_candidate_03.st ---- *)
(* CONTRACT_RULES [{"kind": "hold_until_reset", "output": "tripLatched", "set_input": "runRequest_AND_NOT_pressureValid_OR_pressure_ge_4500", "reset_input": "resetBtn_rising_AND_NOT_runRequest_AND_pressureValid_AND_pressure_le_4200"}] *)
(* ENGINEERING_CONTRACT
   PUB001-PUB004:  Trip activation same-scan when runRequest AND (NOT pressureValid OR pressure >= 4500.0 kPa).
   PUB005:         Hysteresis band 300 kPa: reset clears only when pressure <= 4200.0 (strict <=).
   PUB006-PUB008:  tripLatched holds until resetBtn rising edge + NOT runRequest + pressureValid + pressure <= 4200.0.
   PUB009-PUB011:  currentCauseMask LOW-4 encoding: bit0=xmitter fail, bit1=valve stick(3-consecutive), bit2=excess combustion, bit3=unlocated.
                    Only evaluated when runRequest AND pressureValid AND pressure >= 4500.0 (bits 1/2); bit0 when runRequest AND NOT pressureValid.
                    Not runRequest → mask = 0.
   PUB012-PUB014:  Valve stick counter requires 3 consecutive cycles of (runRequest AND pressureValid AND pressure >= 4500.0 AND outletCmd >= 50 AND outletFeedback <= 10).
                    Any break (feedback OK, pressure < 4500, pressureValid=FALSE, runRequest=FALSE) → counter = 0.
   PUB015-PUB017:  latchedCauseMask accumulates via bitwise OR each scan tripLatched is TRUE (16-bit WORD, max 15, no overflow).
                    Cleared only on legal reset. Reflects full trip history, not a snapshot.
   PUB018-PUB020:  fuelPermit = runRequest AND NOT tripLatched; diagnosticActive = (currentCauseMask <> 0).
   PUB021-PUB023:  Clue encodings: 0=none, 1=xmitter fail, 2=stick only, 4=combustion only, 6=both, 8=unlocated.
   Units: kPa (pressure), t/h (flow), % (valve).
*)
FUNCTION_BLOCK FB
VAR
    prevResetBtn      : BOOL := FALSE;
    prevStickingCond1 : BOOL := FALSE;
    prevStickingCond2 : BOOL := FALSE;
    stickingCount     : INT  := 0;
    local_tripLatched : BOOL := FALSE;
    local_fuelPermit  : BOOL := FALSE;
    local_currentMask : WORD := 16#0000;
    local_latchedMask : WORD := 16#0000;
END_VAR
VAR_TEMP
    resetRising   : BOOL;
    curSticking   : BOOL;
END_VAR

    resetRising := resetBtn AND NOT prevResetBtn;

    IF resetRising AND NOT runRequest AND pressureValid AND (pressure <= 4200.0) THEN
        local_tripLatched := FALSE;
        local_latchedMask := 16#0000;
    ELSIF runRequest AND (NOT pressureValid OR (pressure >= 4500.0)) THEN
        local_tripLatched := TRUE;
    END_IF;

    curSticking := runRequest AND pressureValid AND (pressure >= 4500.0) AND (outletCmd >= 50) AND (outletFeedback <= 10);

    IF curSticking THEN
        IF prevStickingCond1 AND prevStickingCond2 THEN
            stickingCount := 3;
        ELSE
            stickingCount := stickingCount + 1;
            IF stickingCount > 3 THEN
                stickingCount := 3;
            END_IF;
        END_IF;
    ELSE
        stickingCount := 0;
    END_IF;

    local_currentMask := 16#0000;

    IF NOT runRequest THEN
        local_currentMask := 16#0000;
    ELSIF NOT pressureValid THEN
        local_currentMask := 16#0001;
    ELSE
        IF pressure >= 4500.0 THEN
            IF stickingCount >= 3 THEN
                local_currentMask := local_currentMask OR TO_WORD(2);
            END_IF;
            IF (fuelFlow >= 4.0) AND (steamFlow <= 10.0) THEN
                local_currentMask := local_currentMask OR TO_WORD(4);
            END_IF;
            IF (stickingCount < 3) AND NOT ((fuelFlow >= 4.0) AND (steamFlow <= 10.0)) THEN
                local_currentMask := local_currentMask OR TO_WORD(8);
            END_IF;
        END_IF;
    END_IF;

    IF local_tripLatched THEN
        local_latchedMask := local_latchedMask OR local_currentMask;
    END_IF;

    local_fuelPermit := runRequest AND NOT local_tripLatched;

    tripLatched      := local_tripLatched;
    fuelPermit       := local_fuelPermit;
    currentCauseMask := local_currentMask;
    latchedCauseMask := local_latchedMask;
    diagnosticActive := (local_currentMask <> 16#0000);

    prevResetBtn      := resetBtn;
    prevStickingCond2 := prevStickingCond1;
    prevStickingCond1 := curSticking;

END_FUNCTION_BLOCK

(* ---- self-hard-06.raw_candidate_04.st ---- *)
(* CONTRACT_RULES [{"kind": "hold_until_reset", "output": "tripLatched", "set_input": "runRequest_AND_NOT_pressureValid_OR_pressure_ge_4500", "reset_input": "resetBtn_rising_AND_NOT_runRequest_AND_pressureValid_AND_pressure_le_4200"}] *)
(* ENGINEERING_CONTRACT
   PUB001-PUB004:  Trip activation same-scan when runRequest AND (NOT pressureValid OR pressure >= 4500.0 kPa).
   PUB005:         Hysteresis band 300 kPa: reset clears only when pressure <= 4200.0 (strict <=).
   PUB006-PUB008:  tripLatched holds until resetBtn rising edge + NOT runRequest + pressureValid + pressure <= 4200.0.
   PUB009-PUB011:  currentCauseMask LOW-4 encoding: bit0=xmitter fail, bit1=valve stick(3-consecutive), bit2=excess combustion, bit3=unlocated.
                    Only evaluated when runRequest AND pressureValid AND pressure >= 4500.0 (bits 1/2); bit0 when runRequest AND NOT pressureValid.
                    Not runRequest → mask = 0.
   PUB012-PUB014:  Valve stick counter requires 3 consecutive cycles of (runRequest AND pressureValid AND pressure >= 4500.0 AND outletCmd >= 50 AND outletFeedback <= 10).
                    Any break (feedback OK, pressure < 4500, pressureValid=FALSE, runRequest=FALSE) → counter = 0.
   PUB015-PUB017:  latchedCauseMask accumulates via bitwise OR each scan tripLatched is TRUE (16-bit WORD, max 15, no overflow).
                    Cleared only on legal reset. Reflects full trip history, not a snapshot.
   PUB018-PUB020:  fuelPermit = runRequest AND NOT tripLatched; diagnosticActive = (currentCauseMask <> 0).
   PUB021-PUB023:  Clue encodings: 0=none, 1=xmitter fail, 2=stick only, 4=combustion only, 6=both, 8=unlocated.
   Units: kPa (pressure), t/h (flow), % (valve).
*)
FUNCTION_BLOCK FB
VAR
    prevResetBtn      : BOOL := FALSE;
    prevStickingCond1 : BOOL := FALSE;
    prevStickingCond2 : BOOL := FALSE;
    stickingCount     : INT  := 0;
    tmpResetRising    : BOOL := FALSE;
END_VAR
VAR_OUTPUT
    tripLatched       : BOOL;
    fuelPermit        : BOOL;
    currentCauseMask  : WORD;
    latchedCauseMask  : WORD;
    diagnosticActive  : BOOL;
END_VAR

    // Rising-edge detection for reset button (PUB006)
    tmpResetRising := resetBtn AND NOT prevResetBtn;

    // Trip condition: set or clear tripLatched (PUB001-PUB004, S1, S2, S17)
    IF tmpResetRising AND NOT runRequest AND pressureValid AND (pressure <= 4200.0) THEN
        tripLatched := FALSE;
    ELSIF runRequest AND (NOT pressureValid OR (pressure >= 4500.0)) THEN
        tripLatched := TRUE;
    END_IF;

    // Valve sticking: 3 consecutive cycles under valid overpressure (PUB012-PUB014, N10-S11)
    IF runRequest AND pressureValid AND (pressure >= 4500.0) AND (outletCmd >= 50) AND (outletFeedback <= 10) THEN
        IF prevStickingCond1 AND prevStickingCond2 THEN
            stickingCount := 3;
        ELSE
            stickingCount := stickingCount + 1;
            IF stickingCount > 3 THEN
                stickingCount := 3;
            END_IF;
        END_IF;
    ELSE
        stickingCount := 0;
    END_IF;

    // Current cause mask (PUB009-PUB011, S5, S6, S9-S12, N10-S10, N10-S11, N10-S15)
    currentCauseMask := 16#0000;

    IF NOT runRequest THEN
        currentCauseMask := 16#0000;
    ELSIF NOT pressureValid THEN
        currentCauseMask := 16#0001;
    ELSE
        IF pressure >= 4500.0 THEN
            IF stickingCount >= 3 THEN
                currentCauseMask := currentCauseMask OR INT_TO_WORD(2);
            END_IF;
            IF (fuelFlow >= 4.0) AND (steamFlow <= 10.0) THEN
                currentCauseMask := currentCauseMask OR INT_TO_WORD(4);
            END_IF;
            IF (stickingCount < 3) AND NOT ((fuelFlow >= 4.0) AND (steamFlow <= 10.0)) THEN
                currentCauseMask := currentCauseMask OR INT_TO_WORD(8);
            END_IF;
        END_IF;
    END_IF;

    // Latched cause mask accumulation (PUB015-PUB017, S13, N10-S18)
    IF tripLatched AND (currentCauseMask <> 16#0000) THEN
        latchedCauseMask := latchedCauseMask OR currentCauseMask;
    END_IF;

    // Outputs (PUB018-PUB020, S3, N10-S16)
    fuelPermit       := runRequest AND NOT tripLatched;
    diagnosticActive := (currentCauseMask <> 16#0000);

    // State propagation for next scan
    prevResetBtn      := resetBtn;
    prevStickingCond2 := prevStickingCond1;
    prevStickingCond1 := (runRequest AND pressureValid AND (pressure >= 4500.0) AND (outletCmd >= 50) AND (outletFeedback <= 10));

END_FUNCTION_BLOCK

(* ---- self-hard-07.candidate_01.st ---- *)
FUNCTION_BLOCK FB
VAR_INPUT
    mode            : INT;
    resetBtn        : BOOL;
    scanSeconds     : REAL;
    tempSP          : REAL;
    tempPV          : REAL;
    flowPV          : REAL;
    manualFlowSP    : REAL;
    manualValve     : REAL;
END_VAR

VAR_OUTPUT
    flowSP          : REAL;
    valveCommand    : REAL;
    fault           : BOOL;
    normalMode      : BOOL;
END_VAR

VAR
    prevMode            : INT := -1;
    prevResetBtn        : BOOL := FALSE;
    firstScan           : BOOL := TRUE;
    prevFlowSP          : REAL := 0.0;
    prevValveCommand    : REAL := 0.0;
    prevTempSP          : REAL := 0.0;
    prevFlowSP_inner    : REAL := 0.0;
    accT                : REAL := 0.0;  // Outer-loop integrator (t/h)
    accF                : REAL := 0.0;  // Inner-loop integrator (%)
    tmpModeSwitch       : BOOL := FALSE;
END_VAR

(* ENGINEERING_CONTRACT
================================================================================
OUTPUT STATE TABLE (per scan, evaluated in priority order):
--------------------------------------------------------------------------------
| State          | Activation        | Retention    | Reset/Deactivation      |
|----------------|-------------------|--------------|-------------------------|
| fault=TRUE     | mode∉{0,1,2} OR   | Hold (latch) | mode returns to 0/1/2   |
|                | scanSeconds≤0 OR  |              | AND scanSeconds valid   |
|                | scanSeconds>10    |              |                         |
| normalMode=TRUE| Mode stable, no   | Same-scan    | Any mode change, fault, |
|                | fault, no reset   | priority     | or reset rising edge    |
| flowSP         | PI output/bumpless| Hold in most | Reset/fault: manualFlowSP|
|                | transfer per mode | modes        | Switch to 0/1: manualSP |
| valveCommand   | PI output/manual  | Hold on      | Reset/fault: manualValve|
|                | per mode          | switch 0/1/2 | Switch 0/1: prev value  |
--------------------------------------------------------------------------------
CONTROLLER GAINS (per PUB003/PUB004):
  Outer loop (temp→flow): KpT=1.0 (t/h)/℃, KiT=0.2 (t/h)/(℃·s)
  Inner loop (flow→valve): KpF=2.0 %/(t/h), KiF=0.5 %/((t/h)·s)
UNITS/BOUNDARIES (PUB001/PUB002):
  flowSP: 0..50 t/h; valveCommand: 0..100 %
ANTI-WINDUP (PUB006): Back-calculation from clamped output
FIRST-SCAN (PUB049): Outputs preset to manual values, normalMode=FALSE
RESET PRIORITY (PUB051/PUB052/PUB053): Outputs/integrators preset; fault still
  reported based on current mode/scanSeconds
FAULT PRIORITY (PUB051/PUB052/PUB053): Immediate manual-follow, no integration;
  fault reported based on current mode/scanSeconds
================================================================================
*)

(* CONTRACT_RULES [] *)

tmpModeSwitch := (prevMode <> mode);

IF firstScan THEN
    // PUB049: First scan preset
    flowSP := manualFlowSP;
    valveCommand := manualValve;
    firstScan := FALSE;
    RETURN;
END_IF;

// PUB050: Fault detection - mode out of range or scanSeconds invalid
fault := (mode < 0) OR (mode > 2) OR (scanSeconds <= 0.0) OR (scanSeconds > 10.0);

// PUB051/PUB052/PUB053: Reset rising edge takes priority for outputs/integrators
IF resetBtn AND NOT prevResetBtn THEN
    flowSP := manualFlowSP;
    valveCommand := manualValve;
    accT := 0.0;
    accF := 0.0;
    prevResetBtn := TRUE;
    prevMode := mode;
    prevFlowSP := flowSP;
    prevValveCommand := valveCommand;
    prevTempSP := tempSP;
    prevFlowSP_inner := flowSP;
    RETURN;
END_IF;
prevResetBtn := resetBtn;

// PUB052: Fault action - immediate manual-follow, integrator preset
IF fault THEN
    flowSP := manualValve;
    valveCommand := manualValve;
    accT := 0.0;
    accF := 0.0;
    normalMode := FALSE;
    prevMode := mode;
    prevFlowSP := flowSP;
    prevValveCommand := valveCommand;
    prevTempSP := tempSP;
    prevFlowSP_inner := flowSP;
    RETURN;
END_IF;

// PUB054/PUB055/PUB056/PUB057/PUB058: Bumpless transfer on mode switch
IF tmpModeSwitch THEN
    normalMode := FALSE;
    // PUB054/PUB055: Switch to manual(0) or auto(1)
    IF mode = 0 OR mode = 1 THEN
        flowSP := manualFlowSP;
        // PUB057: Valve holds previous value
        valveCommand := prevValveCommand;
    // PUB056/PUB058: Switch to cascade(2)
    ELSIF mode = 2 THEN
        // PUB058: Both outputs hold previous values
        flowSP := prevFlowSP;
        valveCommand := prevValveCommand;
    END_IF;
ELSE
    // Normal operation - PI execution
    normalMode := TRUE;

    CASE mode OF
        0: // PUB059: Manual - both outputs follow manual
            flowSP := manualFlowSP;
            valveCommand := manualValve;

        1: // PUB059: Auto - flow manual, inner PI active
            flowSP := manualFlowSP;
            // Inner loop PI with anti-windup back-calculation
            // eF = flowSP - flowPV; trial = accF + 0.5*eF*scanSeconds
            // valveCommand = LIMIT(0, 2.0*eF + trial, 100)
            // accF = valveCommand - 2.0*eF
            prevFlowSP_inner := flowSP;  // Store for inner-loop back-calculation
            accF := prevValveCommand - 2.0 * (prevFlowSP_inner - prevFlowSP_inner);  // Simplified for auto
            // Re-evaluate with proper flowPV
            accF := prevValveCommand - 2.0 * (prevFlowSP_inner - prevFlowSP_inner);
            accF := prevValveCommand - 2.0 * (prevFlowSP_inner - prevFlowSP_inner);
            // Correct inner loop calculation
            prevFlowSP_inner := flowSP;
            accF := prevValveCommand - 2.0 * (flowSP - flowPV);
            valveCommand := LIMIT(0.0, 2.0 * (flowSP - flowPV) + accF, 100.0);
            accF := valveCommand - 2.0 * (flowSP - flowPV);

        2: // PUB059: Cascade - both PI loops active
            // Outer loop PI (temperature → flow)
            // eT = tempSP - tempPV
            // trial = accT + 0.2*eT*scanSeconds
            // flowSP = LIMIT(0, 1.0*eT + trial, 50)
            // accT = flowSP - 1.0*eT
            accT := prevFlowSP - 1.0 * prevTempSP;
            flowSP := LIMIT(0.0, 1.0 * (tempSP - tempPV) + accT + 0.2 * (tempSP - tempPV) * scanSeconds, 50.0);
            accT := flowSP - 1.0 * (tempSP - tempPV);

            // Inner loop PI (flow → valve) using current flowSP
            // eF = flowSP - flowPV
            // trial = accF + 0.5*eF*scanSeconds
            // valveCommand = LIMIT(0, 2.0*eF + trial, 100)
            // accF = valveCommand - 2.0*eF
            prevFlowSP_inner := prevFlowSP;
            accF := prevValveCommand - 2.0 * (prevFlowSP_inner - prevFlowSP_inner);
            accF := prevValveCommand - 2.0 * (prevFlowSP - flowPV);
            valveCommand := LIMIT(0.0, 2.0 * (flowSP - flowPV) + accF + 0.5 * (flowSP - flowPV) * scanSeconds, 100.0);
            accF := valveCommand - 2.0 * (flowSP - flowPV);
    END_CASE;
END_IF;

// Update state for next scan
prevMode := mode;
prevFlowSP := flowSP;
prevValveCommand := valveCommand;
prevTempSP := tempSP;
prevFlowSP_inner := prevFlowSP_inner;  // Preserve for back-calculation

END_FUNCTION_BLOCK

(* ---- self-hard-07.candidate_02.st ---- *)
FUNCTION_BLOCK FB
VAR_INPUT
    mode            : INT;
    resetBtn        : BOOL;
    scanSeconds     : REAL;
    tempSP          : REAL;
    tempPV          : REAL;
    flowPV          : REAL;
    manualFlowSP    : REAL;
    manualValve     : REAL;
END_VAR

VAR_OUTPUT
    flowSP          : REAL;
    valveCommand    : REAL;
    fault           : BOOL;
    normalMode      : BOOL;
END_VAR

VAR
    prevMode            : INT := -1;
    prevResetBtn        : BOOL := FALSE;
    firstScan           : BOOL := TRUE;
    prevFlowSP          : REAL := 0.0;
    prevValveCommand    : REAL := 0.0;
    prevTempSP          : REAL := 0.0;
    prevFlowSP_inner    : REAL := 0.0;
    accT                : REAL := 0.0;
    accF                : REAL := 0.0;
    tmpModeSwitch       : BOOL := FALSE;
END_VAR

(* ENGINEERING_CONTRACT
================================================================================
OUTPUT STATE TABLE (per scan, evaluated in priority order):
--------------------------------------------------------------------------------
| State          | Activation        | Retention    | Reset/Deactivation      |
|----------------|-------------------|--------------|-------------------------|
| fault=TRUE     | mode∉{0,1,2} OR   | Hold (latch) | mode returns to 0/1/2   |
|                | scanSeconds≤0 OR  |              | AND scanSeconds valid   |
|                | scanSeconds>10    |              |                         |
| normalMode=TRUE| Mode stable, no   | Same-scan    | Any mode change, fault, |
|                | fault, no reset   | priority     | or reset rising edge    |
| flowSP         | PI output/bumpless| Hold in most | Reset/fault: manualFlowSP|
|                | transfer per mode | modes        | Switch to 0/1: manualSP |
| valveCommand   | PI output/manual  | Hold on      | Reset/fault: manualValve|
|                | per mode          | switch 0/1/2 | Switch 0/1: prev value  |
--------------------------------------------------------------------------------
CONTROLLER GAINS (per PUB003/PUB004):
  Outer loop (temp→flow): KpT=1.0 (t/h)/℃, KiT=0.2 (t/h)/(℃·s)
  Inner loop (flow→valve): KpF=2.0 %/(t/h), KiF=0.5 %/((t/h)·s)
UNITS/BOUNDARIES (PUB001/PUB002):
  flowSP: 0..50 t/h; valveCommand: 0..100 %
ANTI-WINDUP (PUB006): Back-calculation from clamped output
FIRST-SCAN (PUB049): Outputs preset to manual values, normalMode=FALSE
RESET PRIORITY (PUB051/PUB052/PUB053): Outputs/integrators preset; fault still
  reported based on current mode/scanSeconds
FAULT PRIORITY (PUB051/PUB052/PUB053): Immediate manual-follow, no integration;
  fault reported based on current mode/scanSeconds
================================================================================
*)

(* CONTRACT_RULES [] *)

tmpModeSwitch := (prevMode <> mode) AND NOT firstScan;

IF firstScan THEN
    // PUB049: First scan preset - also initialize prevMode for correct switch detection
    flowSP := manualFlowSP;
    valveCommand := manualValve;
    prevMode := mode;
    firstScan := FALSE;
    RETURN;
END_IF;

// PUB050: Fault detection - mode out of range or scanSeconds invalid
fault := (mode < 0) OR (mode > 2) OR (scanSeconds <= 0.0) OR (scanSeconds > 10.0);

// PUB051/PUB052/PUB053: Reset rising edge takes priority for outputs/integrators
IF resetBtn AND NOT prevResetBtn THEN
    flowSP := manualFlowSP;
    valveCommand := manualValve;
    accT := 0.0;
    accF := 0.0;
    prevResetBtn := TRUE;
    prevMode := mode;
    prevFlowSP := flowSP;
    prevValveCommand := valveCommand;
    prevTempSP := tempSP;
    prevFlowSP_inner := flowSP;
    RETURN;
END_IF;
prevResetBtn := resetBtn;

// PUB052: Fault action - immediate manual-follow, integrator preset
IF fault THEN
    flowSP := manualFlowSP;
    valveCommand := manualValve;
    accT := 0.0;
    accF := 0.0;
    normalMode := FALSE;
    prevMode := mode;
    prevFlowSP := flowSP;
    prevValveCommand := valveCommand;
    prevTempSP := tempSP;
    prevFlowSP_inner := flowSP;
    RETURN;
END_IF;

// PUB054/PUB055/PUB056/PUB057/PUB058: Bumpless transfer on mode switch
IF tmpModeSwitch THEN
    normalMode := FALSE;
    // PUB054/PUB055: Switch to manual(0) or auto(1)
    IF (mode = 0) OR (mode = 1) THEN
        flowSP := manualFlowSP;
        // PUB057: Valve holds previous value
        valveCommand := prevValveCommand;
    // PUB056/PUB058: Switch to cascade(2)
    ELSIF mode = 2 THEN
        // PUB058: Both outputs hold previous values
        flowSP := prevFlowSP;
        valveCommand := prevValveCommand;
    END_IF;
ELSE
    // Normal operation - PI execution
    normalMode := TRUE;

    CASE mode OF
        0: // PUB059: Manual - both outputs follow manual
            flowSP := manualFlowSP;
            valveCommand := manualValve;

        1: // PUB059: Auto - flow manual, inner PI active
            flowSP := manualFlowSP;
            // Inner loop PI with anti-windup back-calculation
            prevFlowSP_inner := flowSP;
            accF := prevValveCommand - 2.0 * (prevFlowSP_inner - flowPV);
            valveCommand := LIMIT(0.0, 2.0 * (flowSP - flowPV) + accF + 0.5 * (flowSP - flowPV) * scanSeconds, 100.0);
            accF := valveCommand - 2.0 * (flowSP - flowPV);

        2: // PUB059: Cascade - both PI loops active
            // Outer loop PI (temperature → flow)
            accT := prevFlowSP - 1.0 * prevTempSP;
            flowSP := LIMIT(0.0, 1.0 * (tempSP - tempPV) + accT + 0.2 * (tempSP - tempPV) * scanSeconds, 50.0);
            accT := flowSP - 1.0 * (tempSP - tempPV);

            // Inner loop PI (flow → valve) using current flowSP
            prevFlowSP_inner := prevFlowSP;
            accF := prevValveCommand - 2.0 * (prevFlowSP_inner - flowPV);
            valveCommand := LIMIT(0.0, 2.0 * (flowSP - flowPV) + accF + 0.5 * (flowSP - flowPV) * scanSeconds, 100.0);
            accF := valveCommand - 2.0 * (flowSP - flowPV);
    END_CASE;
END_IF;

// Update state for next scan
prevMode := mode;
prevFlowSP := flowSP;
prevValveCommand := valveCommand;
prevTempSP := tempSP;
prevFlowSP_inner := flowSP;

END_FUNCTION_BLOCK

(* ---- self-hard-07.candidate_03.st ---- *)
FUNCTION_BLOCK FB
VAR_INPUT
    mode            : INT;
    resetBtn        : BOOL;
    scanSeconds     : REAL;
    tempSP          : REAL;
    tempPV          : REAL;
    flowPV          : REAL;
    manualFlowSP    : REAL;
    manualValve     : REAL;
END_VAR

VAR_OUTPUT
    flowSP          : REAL;
    valveCommand    : REAL;
    fault           : BOOL;
    normalMode      : BOOL;
END_VAR

VAR
    prevMode            : INT := -1;
    prevResetBtn        : BOOL := FALSE;
    firstScan           : BOOL := TRUE;
    prevFlowSP          : REAL := 0.0;
    prevValveCommand    : REAL := 0.0;
    prevTempSP          : REAL := 0.0;
    prevFlowSP_inner    : REAL := 0.0;
    accT                : REAL := 0.0;
    accF                : REAL := 0.0;
    tmpModeSwitch       : BOOL := FALSE;
END_VAR

(* ENGINEERING_CONTRACT
================================================================================
OUTPUT STATE TABLE (per scan, evaluated in priority order):
--------------------------------------------------------------------------------
| State          | Activation        | Retention    | Reset/Deactivation      |
|----------------|-------------------|--------------|-------------------------|
| fault=TRUE     | mode∉{0,1,2} OR   | Hold (latch) | mode returns to 0/1/2   |
|                | scanSeconds≤0 OR  |              | AND scanSeconds valid   |
|                | scanSeconds>10    |              |                         |
| normalMode=TRUE| Mode stable, no   | Same-scan    | Any mode change, fault, |
|                | fault, no reset   | priority     | or reset rising edge    |
| flowSP         | PI output/bumpless| Hold in most | Reset/fault: manualFlowSP|
|                | transfer per mode | modes        | Switch to 0/1: manualSP |
| valveCommand   | PI output/manual  | Hold on      | Reset/fault: manualValve|
|                | per mode          | switch 0/1/2 | Switch 0/1: prev value  |
--------------------------------------------------------------------------------
CONTROLLER GAINS (per PUB003/PUB004):
  Outer loop (temp→flow): KpT=1.0 (t/h)/℃, KiT=0.2 (t/h)/(℃·s)
  Inner loop (flow→valve): KpF=2.0 %/(t/h), KiF=0.5 %/((t/h)·s)
UNITS/BOUNDARIES (PUB001/PUB002):
  flowSP: 0..50 t/h; valveCommand: 0..100 %
ANTI-WINDUP (PUB006): Back-calculation from clamped output
FIRST-SCAN (PUB049): Outputs preset to manual values, normalMode=FALSE
RESET PRIORITY (PUB051/PUB052/PUB053): Outputs/integrators preset; fault still
  reported based on current mode/scanSeconds
FAULT PRIORITY (PUB051/PUB052/PUB053): Immediate manual-follow, no integration;
  fault reported based on current mode/scanSeconds
================================================================================
*)

(* CONTRACT_RULES [] *)

tmpModeSwitch := (prevMode <> mode) AND NOT firstScan;

IF firstScan THEN
    flowSP := manualFlowSP;
    valveCommand := manualValve;
    prevMode := mode;
    firstScan := FALSE;
END_IF;

// PUB050: Fault detection - mode out of range or scanSeconds invalid
fault := (mode < 0) OR (mode > 2) OR (scanSeconds <= 0.0) OR (scanSeconds > 10.0);

// PUB051/PUB052/PUB053: Reset rising edge takes priority for outputs/integrators
IF resetBtn AND NOT prevResetBtn THEN
    flowSP := manualFlowSP;
    valveCommand := manualValve;
    accT := 0.0;
    accF := 0.0;
    prevResetBtn := TRUE;
    prevMode := mode;
    prevFlowSP := flowSP;
    prevValveCommand := valveCommand;
    prevTempSP := tempSP;
    prevFlowSP_inner := flowSP;
    RETURN;
END_IF;
prevResetBtn := resetBtn;

// PUB052: Fault action - immediate manual-follow, integrator preset
IF fault THEN
    flowSP := manualFlowSP;
    valveCommand := manualValve;
    accT := 0.0;
    accF := 0.0;
    normalMode := FALSE;
    prevMode := mode;
    prevFlowSP := flowSP;
    prevValveCommand := valveCommand;
    prevTempSP := tempSP;
    prevFlowSP_inner := flowSP;
    RETURN;
END_IF;

// PUB054/PUB055/PUB056/PUB057/PUB058: Bumpless transfer on mode switch
IF tmpModeSwitch THEN
    normalMode := FALSE;
    // PUB054/PUB055: Switch to manual(0) or auto(1)
    IF (mode = 0) OR (mode = 1) THEN
        flowSP := manualFlowSP;
        // PUB057: Valve holds previous value
        valveCommand := prevValveCommand;
    // PUB056/PUB058: Switch to cascade(2)
    ELSIF mode = 2 THEN
        // PUB058: Both outputs hold previous values
        flowSP := prevFlowSP;
        valveCommand := prevValveCommand;
    END_IF;
ELSE
    // Normal operation - PI execution
    normalMode := TRUE;

    CASE mode OF
        0: // PUB059: Manual - both outputs follow manual
            flowSP := manualFlowSP;
            valveCommand := manualValve;

        1: // PUB059: Auto - flow manual, inner PI active
            flowSP := manualFlowSP;
            // Inner loop PI with anti-windup back-calculation
            accF := prevValveCommand - 2.0 * (prevFlowSP_inner - flowPV);
            valveCommand := LIMIT(0.0, 2.0 * (flowSP - flowPV) + accF + 0.5 * (flowSP - flowPV) * scanSeconds, 100.0);
            accF := valveCommand - 2.0 * (flowSP - flowPV);

        2: // PUB059: Cascade - both PI loops active
            // Outer loop PI (temperature → flow)
            accT := prevFlowSP - 1.0 * prevTempSP;
            flowSP := LIMIT(0.0, 1.0 * (tempSP - tempPV) + accT + 0.2 * (tempSP - tempPV) * scanSeconds, 50.0);
            accT := flowSP - 1.0 * (tempSP - tempPV);

            // Inner loop PI (flow → valve) using current flowSP
            accF := prevValveCommand - 2.0 * (prevFlowSP_inner - flowPV);
            valveCommand := LIMIT(0.0, 2.0 * (flowSP - flowPV) + accF + 0.5 * (flowSP - flowPV) * scanSeconds, 100.0);
            accF := valveCommand - 2.0 * (flowSP - flowPV);
    END_CASE;
END_IF;

// Update state for next scan
prevMode := mode;
prevFlowSP := flowSP;
prevValveCommand := valveCommand;
prevTempSP := tempSP;
prevFlowSP_inner := flowSP;

END_FUNCTION_BLOCK

(* ---- self-hard-07.raw_candidate_01.st ---- *)
FUNCTION_BLOCK FB
VAR_INPUT
    mode            : INT;
    resetBtn        : BOOL;
    scanSeconds     : REAL;
    tempSP          : REAL;
    tempPV          : REAL;
    flowPV          : REAL;
    manualFlowSP    : REAL;
    manualValve     : REAL;
END_VAR

VAR_OUTPUT
    flowSP          : REAL;
    valveCommand    : REAL;
    fault           : BOOL;
    normalMode      : BOOL;
END_VAR

VAR
    prevMode            : INT := -1;
    prevResetBtn        : BOOL := FALSE;
    firstScan           : BOOL := TRUE;
    prevFlowSP          : REAL := 0.0;
    prevValveCommand    : REAL := 0.0;
    prevTempSP          : REAL := 0.0;
    prevFlowSP_inner    : REAL := 0.0;
    accT                : REAL := 0.0;  // Outer-loop integrator (t/h)
    accF                : REAL := 0.0;  // Inner-loop integrator (%)
    tmpModeSwitch       : BOOL := FALSE;
END_VAR

(* ENGINEERING_CONTRACT
================================================================================
OUTPUT STATE TABLE (per scan, evaluated in priority order):
--------------------------------------------------------------------------------
| State          | Activation        | Retention    | Reset/Deactivation      |
|----------------|-------------------|--------------|-------------------------|
| fault=TRUE     | mode∉{0,1,2} OR   | Hold (latch) | mode returns to 0/1/2   |
|                | scanSeconds≤0 OR  |              | AND scanSeconds valid   |
|                | scanSeconds>10    |              |                         |
| normalMode=TRUE| Mode stable, no   | Same-scan    | Any mode change, fault, |
|                | fault, no reset   | priority     | or reset rising edge    |
| flowSP         | PI output/bumpless| Hold in most | Reset/fault: manualFlowSP|
|                | transfer per mode | modes        | Switch to 0/1: manualSP |
| valveCommand   | PI output/manual  | Hold on      | Reset/fault: manualValve|
|                | per mode          | switch 0/1/2 | Switch 0/1: prev value  |
--------------------------------------------------------------------------------
CONTROLLER GAINS (per PUB003/PUB004):
  Outer loop (temp→flow): KpT=1.0 (t/h)/℃, KiT=0.2 (t/h)/(℃·s)
  Inner loop (flow→valve): KpF=2.0 %/(t/h), KiF=0.5 %/((t/h)·s)
UNITS/BOUNDARIES (PUB001/PUB002):
  flowSP: 0..50 t/h; valveCommand: 0..100 %
ANTI-WINDUP (PUB006): Back-calculation from clamped output
FIRST-SCAN (PUB049): Outputs preset to manual values, normalMode=FALSE
RESET PRIORITY (PUB051/PUB052/PUB053): Outputs/integrators preset; fault still
  reported based on current mode/scanSeconds
FAULT PRIORITY (PUB051/PUB052/PUB053): Immediate manual-follow, no integration;
  fault reported based on current mode/scanSeconds
================================================================================
*)

(* CONTRACT_RULES [] *)

tmpModeSwitch := (prevMode <> mode);

IF firstScan THEN
    // PUB049: First scan preset
    flowSP := manualFlowSP;
    valveCommand := manualValve;
    firstScan := FALSE;
    RETURN;
END_IF;

// PUB050: Fault detection - mode out of range or scanSeconds invalid
fault := (mode < 0) OR (mode > 2) OR (scanSeconds <= 0.0) OR (scanSeconds > 10.0);

// PUB051/PUB052/PUB053: Reset rising edge takes priority for outputs/integrators
IF resetBtn AND NOT prevResetBtn THEN
    flowSP := manualFlowSP;
    valveCommand := manualValve;
    accT := 0.0;
    accF := 0.0;
    prevResetBtn := TRUE;
    prevMode := mode;
    prevFlowSP := flowSP;
    prevValveCommand := valveCommand;
    prevTempSP := tempSP;
    prevFlowSP_inner := flowSP;
    RETURN;
END_IF;
prevResetBtn := resetBtn;

// PUB052: Fault action - immediate manual-follow, integrator preset
IF fault THEN
    flowSP := manualValve;
    valveCommand := manualValve;
    accT := 0.0;
    accF := 0.0;
    normalMode := FALSE;
    prevMode := mode;
    prevFlowSP := flowSP;
    prevValveCommand := valveCommand;
    prevTempSP := tempSP;
    prevFlowSP_inner := flowSP;
    RETURN;
END_IF;

// PUB054/PUB055/PUB056/PUB057/PUB058: Bumpless transfer on mode switch
IF tmpModeSwitch THEN
    normalMode := FALSE;
    // PUB054/PUB055: Switch to manual(0) or auto(1)
    IF mode = 0 OR mode = 1 THEN
        flowSP := manualFlowSP;
        // PUB057: Valve holds previous value
        valveCommand := prevValveCommand;
    // PUB056/PUB058: Switch to cascade(2)
    ELSIF mode = 2 THEN
        // PUB058: Both outputs hold previous values
        flowSP := prevFlowSP;
        valveCommand := prevValveCommand;
    END_IF;
ELSE
    // Normal operation - PI execution
    normalMode := TRUE;

    CASE mode OF
        0: // PUB059: Manual - both outputs follow manual
            flowSP := manualFlowSP;
            valveCommand := manualValve;

        1: // PUB059: Auto - flow manual, inner PI active
            flowSP := manualFlowSP;
            // Inner loop PI with anti-windup back-calculation
            // eF = flowSP - flowPV; trial = accF + 0.5*eF*scanSeconds
            // valveCommand = LIMIT(0, 2.0*eF + trial, 100)
            // accF = valveCommand - 2.0*eF
            prevFlowSP_inner := flowSP;  // Store for inner-loop back-calculation
            accF := prevValveCommand - 2.0 * (prevFlowSP_inner - prevFlowSP_inner);  // Simplified for auto
            // Re-evaluate with proper flowPV
            accF := prevValveCommand - 2.0 * (prevFlowSP_inner - prevFlowSP_inner);
            accF := prevValveCommand - 2.0 * (prevFlowSP_inner - prevFlowSP_inner);
            // Correct inner loop calculation
            prevFlowSP_inner := flowSP;
            accF := prevValveCommand - 2.0 * (flowSP - flowPV);
            valveCommand := LIMIT(0.0, 2.0 * (flowSP - flowPV) + accF, 100.0);
            accF := valveCommand - 2.0 * (flowSP - flowPV);

        2: // PUB059: Cascade - both PI loops active
            // Outer loop PI (temperature → flow)
            // eT = tempSP - tempPV
            // trial = accT + 0.2*eT*scanSeconds
            // flowSP = LIMIT(0, 1.0*eT + trial, 50)
            // accT = flowSP - 1.0*eT
            accT := prevFlowSP - 1.0 * prevTempSP;
            flowSP := LIMIT(0.0, 1.0 * (tempSP - tempPV) + accT + 0.2 * (tempSP - tempPV) * scanSeconds, 50.0);
            accT := flowSP - 1.0 * (tempSP - tempPV);

            // Inner loop PI (flow → valve) using current flowSP
            // eF = flowSP - flowPV
            // trial = accF + 0.5*eF*scanSeconds
            // valveCommand = LIMIT(0, 2.0*eF + trial, 100)
            // accF = valveCommand - 2.0*eF
            prevFlowSP_inner := prevFlowSP;
            accF := prevValveCommand - 2.0 * (prevFlowSP_inner - prevFlowSP_inner);
            accF := prevValveCommand - 2.0 * (prevFlowSP - flowPV);
            valveCommand := LIMIT(0.0, 2.0 * (flowSP - flowPV) + accF + 0.5 * (flowSP - flowPV) * scanSeconds, 100.0);
            accF := valveCommand - 2.0 * (flowSP - flowPV);
    END_CASE;
END_IF;

// Update state for next scan
prevMode := mode;
prevFlowSP := flowSP;
prevValveCommand := valveCommand;
prevTempSP := tempSP;
prevFlowSP_inner := prevFlowSP_inner;  // Preserve for back-calculation

END_FUNCTION_BLOCK

(* ---- self-hard-07.raw_candidate_02.st ---- *)
FUNCTION_BLOCK FB
VAR_INPUT
    mode            : INT;
    resetBtn        : BOOL;
    scanSeconds     : REAL;
    tempSP          : REAL;
    tempPV          : REAL;
    flowPV          : REAL;
    manualFlowSP    : REAL;
    manualValve     : REAL;
END_VAR

VAR_OUTPUT
    flowSP          : REAL;
    valveCommand    : REAL;
    fault           : BOOL;
    normalMode      : BOOL;
END_VAR

VAR
    prevMode            : INT := -1;
    prevResetBtn        : BOOL := FALSE;
    firstScan           : BOOL := TRUE;
    prevFlowSP          : REAL := 0.0;
    prevValveCommand    : REAL := 0.0;
    prevTempSP          : REAL := 0.0;
    prevFlowSP_inner    : REAL := 0.0;
    accT                : REAL := 0.0;
    accF                : REAL := 0.0;
    tmpModeSwitch       : BOOL := FALSE;
END_VAR

(* ENGINEERING_CONTRACT
================================================================================
OUTPUT STATE TABLE (per scan, evaluated in priority order):
--------------------------------------------------------------------------------
| State          | Activation        | Retention    | Reset/Deactivation      |
|----------------|-------------------|--------------|-------------------------|
| fault=TRUE     | mode∉{0,1,2} OR   | Hold (latch) | mode returns to 0/1/2   |
|                | scanSeconds≤0 OR  |              | AND scanSeconds valid   |
|                | scanSeconds>10    |              |                         |
| normalMode=TRUE| Mode stable, no   | Same-scan    | Any mode change, fault, |
|                | fault, no reset   | priority     | or reset rising edge    |
| flowSP         | PI output/bumpless| Hold in most | Reset/fault: manualFlowSP|
|                | transfer per mode | modes        | Switch to 0/1: manualSP |
| valveCommand   | PI output/manual  | Hold on      | Reset/fault: manualValve|
|                | per mode          | switch 0/1/2 | Switch 0/1: prev value  |
--------------------------------------------------------------------------------
CONTROLLER GAINS (per PUB003/PUB004):
  Outer loop (temp→flow): KpT=1.0 (t/h)/℃, KiT=0.2 (t/h)/(℃·s)
  Inner loop (flow→valve): KpF=2.0 %/(t/h), KiF=0.5 %/((t/h)·s)
UNITS/BOUNDARIES (PUB001/PUB002):
  flowSP: 0..50 t/h; valveCommand: 0..100 %
ANTI-WINDUP (PUB006): Back-calculation from clamped output
FIRST-SCAN (PUB049): Outputs preset to manual values, normalMode=FALSE
RESET PRIORITY (PUB051/PUB052/PUB053): Outputs/integrators preset; fault still
  reported based on current mode/scanSeconds
FAULT PRIORITY (PUB051/PUB052/PUB053): Immediate manual-follow, no integration;
  fault reported based on current mode/scanSeconds
================================================================================
*)

(* CONTRACT_RULES [] *)

tmpModeSwitch := (prevMode <> mode) AND NOT firstScan;

IF firstScan THEN
    // PUB049: First scan preset - also initialize prevMode for correct switch detection
    flowSP := manualFlowSP;
    valveCommand := manualValve;
    prevMode := mode;
    firstScan := FALSE;
    RETURN;
END_IF;

// PUB050: Fault detection - mode out of range or scanSeconds invalid
fault := (mode < 0) OR (mode > 2) OR (scanSeconds <= 0.0) OR (scanSeconds > 10.0);

// PUB051/PUB052/PUB053: Reset rising edge takes priority for outputs/integrators
IF resetBtn AND NOT prevResetBtn THEN
    flowSP := manualFlowSP;
    valveCommand := manualValve;
    accT := 0.0;
    accF := 0.0;
    prevResetBtn := TRUE;
    prevMode := mode;
    prevFlowSP := flowSP;
    prevValveCommand := valveCommand;
    prevTempSP := tempSP;
    prevFlowSP_inner := flowSP;
    RETURN;
END_IF;
prevResetBtn := resetBtn;

// PUB052: Fault action - immediate manual-follow, integrator preset
IF fault THEN
    flowSP := manualFlowSP;
    valveCommand := manualValve;
    accT := 0.0;
    accF := 0.0;
    normalMode := FALSE;
    prevMode := mode;
    prevFlowSP := flowSP;
    prevValveCommand := valveCommand;
    prevTempSP := tempSP;
    prevFlowSP_inner := flowSP;
    RETURN;
END_IF;

// PUB054/PUB055/PUB056/PUB057/PUB058: Bumpless transfer on mode switch
IF tmpModeSwitch THEN
    normalMode := FALSE;
    // PUB054/PUB055: Switch to manual(0) or auto(1)
    IF (mode = 0) OR (mode = 1) THEN
        flowSP := manualFlowSP;
        // PUB057: Valve holds previous value
        valveCommand := prevValveCommand;
    // PUB056/PUB058: Switch to cascade(2)
    ELSIF mode = 2 THEN
        // PUB058: Both outputs hold previous values
        flowSP := prevFlowSP;
        valveCommand := prevValveCommand;
    END_IF;
ELSE
    // Normal operation - PI execution
    normalMode := TRUE;

    CASE mode OF
        0: // PUB059: Manual - both outputs follow manual
            flowSP := manualFlowSP;
            valveCommand := manualValve;

        1: // PUB059: Auto - flow manual, inner PI active
            flowSP := manualFlowSP;
            // Inner loop PI with anti-windup back-calculation
            prevFlowSP_inner := flowSP;
            accF := prevValveCommand - 2.0 * (prevFlowSP_inner - flowPV);
            valveCommand := LIMIT(0.0, 2.0 * (flowSP - flowPV) + accF + 0.5 * (flowSP - flowPV) * scanSeconds, 100.0);
            accF := valveCommand - 2.0 * (flowSP - flowPV);

        2: // PUB059: Cascade - both PI loops active
            // Outer loop PI (temperature → flow)
            accT := prevFlowSP - 1.0 * prevTempSP;
            flowSP := LIMIT(0.0, 1.0 * (tempSP - tempPV) + accT + 0.2 * (tempSP - tempPV) * scanSeconds, 50.0);
            accT := flowSP - 1.0 * (tempSP - tempPV);

            // Inner loop PI (flow → valve) using current flowSP
            prevFlowSP_inner := prevFlowSP;
            accF := prevValveCommand - 2.0 * (prevFlowSP_inner - flowPV);
            valveCommand := LIMIT(0.0, 2.0 * (flowSP - flowPV) + accF + 0.5 * (flowSP - flowPV) * scanSeconds, 100.0);
            accF := valveCommand - 2.0 * (flowSP - flowPV);
    END_CASE;
END_IF;

// Update state for next scan
prevMode := mode;
prevFlowSP := flowSP;
prevValveCommand := valveCommand;
prevTempSP := tempSP;
prevFlowSP_inner := flowSP;

END_FUNCTION_BLOCK

(* ---- self-hard-07.raw_candidate_03.st ---- *)
FUNCTION_BLOCK FB
VAR_INPUT
    mode            : INT;
    resetBtn        : BOOL;
    scanSeconds     : REAL;
    tempSP          : REAL;
    tempPV          : REAL;
    flowPV          : REAL;
    manualFlowSP    : REAL;
    manualValve     : REAL;
END_VAR

VAR_OUTPUT
    flowSP          : REAL;
    valveCommand    : REAL;
    fault           : BOOL;
    normalMode      : BOOL;
END_VAR

VAR
    prevMode            : INT := -1;
    prevResetBtn        : BOOL := FALSE;
    firstScan           : BOOL := TRUE;
    prevFlowSP          : REAL := 0.0;
    prevValveCommand    : REAL := 0.0;
    prevTempSP          : REAL := 0.0;
    prevFlowSP_inner    : REAL := 0.0;
    accT                : REAL := 0.0;
    accF                : REAL := 0.0;
    tmpModeSwitch       : BOOL := FALSE;
END_VAR

(* ENGINEERING_CONTRACT
================================================================================
OUTPUT STATE TABLE (per scan, evaluated in priority order):
--------------------------------------------------------------------------------
| State          | Activation        | Retention    | Reset/Deactivation      |
|----------------|-------------------|--------------|-------------------------|
| fault=TRUE     | mode∉{0,1,2} OR   | Hold (latch) | mode returns to 0/1/2   |
|                | scanSeconds≤0 OR  |              | AND scanSeconds valid   |
|                | scanSeconds>10    |              |                         |
| normalMode=TRUE| Mode stable, no   | Same-scan    | Any mode change, fault, |
|                | fault, no reset   | priority     | or reset rising edge    |
| flowSP         | PI output/bumpless| Hold in most | Reset/fault: manualFlowSP|
|                | transfer per mode | modes        | Switch to 0/1: manualSP |
| valveCommand   | PI output/manual  | Hold on      | Reset/fault: manualValve|
|                | per mode          | switch 0/1/2 | Switch 0/1: prev value  |
--------------------------------------------------------------------------------
CONTROLLER GAINS (per PUB003/PUB004):
  Outer loop (temp→flow): KpT=1.0 (t/h)/℃, KiT=0.2 (t/h)/(℃·s)
  Inner loop (flow→valve): KpF=2.0 %/(t/h), KiF=0.5 %/((t/h)·s)
UNITS/BOUNDARIES (PUB001/PUB002):
  flowSP: 0..50 t/h; valveCommand: 0..100 %
ANTI-WINDUP (PUB006): Back-calculation from clamped output
FIRST-SCAN (PUB049): Outputs preset to manual values, normalMode=FALSE
RESET PRIORITY (PUB051/PUB052/PUB053): Outputs/integrators preset; fault still
  reported based on current mode/scanSeconds
FAULT PRIORITY (PUB051/PUB052/PUB053): Immediate manual-follow, no integration;
  fault reported based on current mode/scanSeconds
================================================================================
*)

(* CONTRACT_RULES [] *)

tmpModeSwitch := (prevMode <> mode) AND NOT firstScan;

IF firstScan THEN
    flowSP := manualFlowSP;
    valveCommand := manualValve;
    prevMode := mode;
    firstScan := FALSE;
END_IF;

// PUB050: Fault detection - mode out of range or scanSeconds invalid
fault := (mode < 0) OR (mode > 2) OR (scanSeconds <= 0.0) OR (scanSeconds > 10.0);

// PUB051/PUB052/PUB053: Reset rising edge takes priority for outputs/integrators
IF resetBtn AND NOT prevResetBtn THEN
    flowSP := manualFlowSP;
    valveCommand := manualValve;
    accT := 0.0;
    accF := 0.0;
    prevResetBtn := TRUE;
    prevMode := mode;
    prevFlowSP := flowSP;
    prevValveCommand := valveCommand;
    prevTempSP := tempSP;
    prevFlowSP_inner := flowSP;
    RETURN;
END_IF;
prevResetBtn := resetBtn;

// PUB052: Fault action - immediate manual-follow, integrator preset
IF fault THEN
    flowSP := manualFlowSP;
    valveCommand := manualValve;
    accT := 0.0;
    accF := 0.0;
    normalMode := FALSE;
    prevMode := mode;
    prevFlowSP := flowSP;
    prevValveCommand := valveCommand;
    prevTempSP := tempSP;
    prevFlowSP_inner := flowSP;
    RETURN;
END_IF;

// PUB054/PUB055/PUB056/PUB057/PUB058: Bumpless transfer on mode switch
IF tmpModeSwitch THEN
    normalMode := FALSE;
    // PUB054/PUB055: Switch to manual(0) or auto(1)
    IF (mode = 0) OR (mode = 1) THEN
        flowSP := manualFlowSP;
        // PUB057: Valve holds previous value
        valveCommand := prevValveCommand;
    // PUB056/PUB058: Switch to cascade(2)
    ELSIF mode = 2 THEN
        // PUB058: Both outputs hold previous values
        flowSP := prevFlowSP;
        valveCommand := prevValveCommand;
    END_IF;
ELSE
    // Normal operation - PI execution
    normalMode := TRUE;

    CASE mode OF
        0: // PUB059: Manual - both outputs follow manual
            flowSP := manualFlowSP;
            valveCommand := manualValve;

        1: // PUB059: Auto - flow manual, inner PI active
            flowSP := manualFlowSP;
            // Inner loop PI with anti-windup back-calculation
            accF := prevValveCommand - 2.0 * (prevFlowSP_inner - flowPV);
            valveCommand := LIMIT(0.0, 2.0 * (flowSP - flowPV) + accF + 0.5 * (flowSP - flowPV) * scanSeconds, 100.0);
            accF := valveCommand - 2.0 * (flowSP - flowPV);

        2: // PUB059: Cascade - both PI loops active
            // Outer loop PI (temperature → flow)
            accT := prevFlowSP - 1.0 * prevTempSP;
            flowSP := LIMIT(0.0, 1.0 * (tempSP - tempPV) + accT + 0.2 * (tempSP - tempPV) * scanSeconds, 50.0);
            accT := flowSP - 1.0 * (tempSP - tempPV);

            // Inner loop PI (flow → valve) using current flowSP
            accF := prevValveCommand - 2.0 * (prevFlowSP_inner - flowPV);
            valveCommand := LIMIT(0.0, 2.0 * (flowSP - flowPV) + accF + 0.5 * (flowSP - flowPV) * scanSeconds, 100.0);
            accF := valveCommand - 2.0 * (flowSP - flowPV);
    END_CASE;
END_IF;

// Update state for next scan
prevMode := mode;
prevFlowSP := flowSP;
prevValveCommand := valveCommand;
prevTempSP := tempSP;
prevFlowSP_inner := flowSP;

END_FUNCTION_BLOCK

(* ---- self-medium-01.candidate_01.st ---- *)
(* ENGINEERING_CONTRACT *)
(*
  PUB002/PUB005: valid=FALSE → loadedID:=0, valid=TRUE → loadedID:=recipe[selSlot].recipeID
  PUB006: loadCmd rising-edge triggers one-shot load; level-hold does NOT reload
  PUB007: running=TRUE blocks load, loadedID retains previous value
  PUB008: slot out-of-range [1..8] → valid=FALSE, loadedID unchanged; no array OOB access
  PUB009: validation is conjunction: recipeID<>0 AND totalRatio∈[99.0,101.0] AND temperature∈[30.0,180.0]
  Timing: state retention via VAR (static across scans); first-scan prev_* = FALSE (IEC default)
  S1: !running & rising(loadCmd) & valid-slot & empty-slot → valid=FALSE & loadedID=0
  S4/N10-S4: running → loadedID=prev(loadedID) (includes first production entry)
  N10-S9: !running & !rising(loadCmd) → both outputs retain prev value
*)
(* CONTRACT_RULES [] *)

FUNCTION_BLOCK FB
VAR_INPUT
    recipe      : ARRAY[1..8] OF ST_Recipe;
    selSlot     : INT;
    loadCmd     : BOOL;
    running     : BOOL;
END_VAR
VAR_OUTPUT
    valid       : BOOL;
    loadedID    : INT;
END_VAR
VAR
    tmp_loadTrig  : R_TRIG;
    tmp_prevRunning : BOOL := FALSE;
END_VAR

tmp_loadTrig(CLK := loadCmd);

IF tmp_loadTrig.Q AND NOT running THEN
    IF (selSlot >= 1) AND (selSlot <= 8) THEN
        IF (recipe[selSlot].recipeID <> 0) AND
           (recipe[selSlot].totalRatio >= 99.0) AND (recipe[selSlot].totalRatio <= 101.0) AND
           (recipe[selSlot].temperature >= 30.0) AND (recipe[selSlot].temperature <= 180.0) THEN
            valid    := TRUE;
            loadedID := recipe[selSlot].recipeID;
        ELSE
            valid    := FALSE;
            loadedID := 0;
        END_IF;
    ELSE
        valid    := FALSE;
    END_IF;
ELSIF running THEN
    loadedID := loadedID;
END_IF;

tmp_prevRunning := running;

(* ---- self-medium-01.candidate_02.st ---- *)
(* ENGINEERING_CONTRACT *)
(*
  PUB002/PUB005: valid=FALSE → loadedID:=0, valid=TRUE → loadedID:=recipe[selSlot].recipeID
  PUB006: loadCmd rising-edge triggers one-shot load; level-hold does NOT reload
  PUB007: running=TRUE blocks load, loadedID retains previous value
  PUB008: slot out-of-range [1..8] → valid=FALSE, loadedID unchanged; no array OOB access
  PUB009: validation is conjunction: recipeID<>0 AND totalRatio∈[99.0,101.0] AND temperature∈[30.0,180.0]
  Timing: state retention via VAR (static across scans); first-scan prev_* = FALSE (IEC default)
  S1: !running & rising(loadCmd) & valid-slot & empty-slot → valid=FALSE & loadedID=0
  S4/N10-S4: running → loadedID=prev(loadedID) (includes first production entry)
  N10-S9: !running & !rising(loadCmd) → both outputs retain prev value
*)
(* CONTRACT_RULES [] *)

FUNCTION_BLOCK FB
VAR_INPUT
    recipe      : ARRAY[1..8] OF ST_Recipe;
    selSlot     : INT;
    loadCmd     : BOOL;
    running     : BOOL;
END_VAR
VAR_OUTPUT
    valid       : BOOL;
    loadedID    : INT;
END_VAR
VAR
    tmp_loadTrig  : R_TRIG;
    tmp_prevRunning : BOOL := FALSE;
END_VAR

tmp_loadTrig(CLK := loadCmd);

IF tmp_loadTrig.Q AND NOT running THEN
    IF (selSlot >= 1) AND (selSlot <= 8) THEN
        IF (recipe[selSlot].recipeID <> 0) AND
           (recipe[selSlot].totalRatio >= 99.0) AND (recipe[selSlot].totalRatio <= 101.0) AND
           (recipe[selSlot].temperature >= 30.0) AND (recipe[selSlot].temperature <= 180.0) THEN
            valid    := TRUE;
            loadedID := recipe[selSlot].recipeID;
        ELSE
            valid    := FALSE;
            loadedID := 0;
        END_IF;
    ELSE
        valid    := FALSE;
    END_IF;
ELSIF running THEN
    loadedID := loadedID;
END_IF;

tmp_prevRunning := running;
END_FUNCTION_BLOCK
